// TwinCAT 3 PLC project PLC
// Title: ReMeat003
// Company: Total Control
// Author: Vadim Nagdimaev
// ProjectVersion: 0.0.1
// Description: SLD Line
// ProgramVersion: 3.1.4026.27
// libraries:
//   Tc2_SerialCom, * (Beckhoff Automation GmbH)
//   Tc2_Standard, * (Beckhoff Automation GmbH)
//   Tc2_SUPS, * (Beckhoff Automation GmbH)
//   Tc2_System, * (Beckhoff Automation GmbH)
//   Tc2_Utilities, * (Beckhoff Automation GmbH)
//   Tc3_Module, * (Beckhoff Automation GmbH)
//   Util, * (System)
//   VisuDialogs, * (System)
//   BASIC,3.31,OSCAT
// project tree:
//   00 Library/00-General/ CheckBounds.TcPOU
//   00 Library/00-General/TimeAndDate/ FUN_DeltaTime.TcPOU (excluded from build), GVL_Time_12.TcGVL, prg_RealClock.TcPOU
//   00 Library/00-General/UserGroup/ E_userGroup.TcDUT, prg_User.TcPOU
//   00 Library/01 Piston/ E_ErrorPiton.TcDUT, E_PistonDefault_CMD.TcDUT, E_Piston_Recipe_State.TcDUT, E_Piston_State.TcDUT, FB_Piston.TcPOU, FB_Piston_U_L.TcPOU, ST_Piston.TcDUT, ST_Piston_SelectionList.TcDUT, ST_Piston_Setting_Param.TcDUT, ST_Piston_U_L.TcDUT, TextList_Piston_Recipe_State.TcTLO, TextList_Piston_Recipe_State_CloseOpen.TcTLO, TextList_Piston_Recipe_State_DownUp.TcTLO, TextList_Piston_Recipe_State_InOut.TcTLO, TextList_Piston_Recipe_State_OnOff.TcTLO, TextList_Piston_Recipe_State_OpenClose.TcTLO, TextList_Piston_Recipe_State_UpDown.TcTLO
//   00 Library/01 Piston/VISU/ vis_Piston_Control1.TcVIS, vis_Piston_Control1_Compact.TcVIS, vis_Piston_Control2_CloseOpen.TcVIS, vis_Piston_Control2_OpenClose.TcVIS, vis_Piston_Select.TcVIS (excluded from build), vis_Piston_Select_1.TcVIS (excluded from build), vis_Piston_Setting_Table.TcVIS, vis_Piston_Times.TcVIS
//   00 Library/02 Pump/02.1 Dosing Pump/ FB_DosingPump.TcPOU
//   00 Library/02 Pump/ ControlWordStruct.TcDUT, FB_Pump.TcPOU, StatusWordStruct.TcDUT, ST_Pump.TcDUT
//   00 Library/03 SFC/ FB_SFC_Cycle.TcPOU, FB_SFC_Template.TcPOU, ITF_FB_SFC_Cycle.TcIO, ST_SFC.TcDUT, vis_Cycle_Control.TcVIS, vis_Cycle_Control_1.TcVIS, vis_Cycle_Panel.TcVIS
//   00 Library/04 Recipe/ E_Recipe_Root_Folder.TcDUT, FB_Recipe.TcPOU, FB_Recipe_Vizu.TcVIS, GVL_Recipe.TcGVL, ST_Recipe.TcDUT, TextList_RecipeRootFolder.TcTLO
//   00 Library/04 Recipe/OLD/ prg_RecipeManager.TcPOU, vis_RecipeControl_v01.TcVIS, vis_RecipeTest.TcVIS
//   00 Library/04-Messages/DUTs/Errors/ E_ErrorFormat.TcDUT, ST_Error.TcDUT, ST_Mess_Logger.TcDUT
//   00 Library/04-Messages/DUTs/ stMessageFormat.TcDUT
//   00 Library/04-Messages/ FB_PrintErrMessageByID.TcPOU, FB_PrintErrMessageByID_SFC_Cycle.TcPOU, FB_PrintErrMessageByID_ST_Cycle.TcPOU, FUN_Write_Line_To_History.TcPOU, F_iFB_Num_sFB_Num.TcPOU, GVL_CycleMessages.TcGVL
//   00 Library/05 Safety/ FB_TwinSAFE.TcPOU, GVL_Safety.TcGVL, prg_Safety.TcPOU, ST_ES_PB.TcDUT, ST_SafeOut_PlcIn.TcDUT, ST_SafeIn_PlcOut.TcDUT, Vis_ES_PB.TcVIS
//   00 Library/05 Safety/TwinSAFE/ e_DualChanal.TcDUT, TwinSafeOut_PlcIn.TcDUT, TwinSafeIn_PlcOut.TcDUT
//   00 Library/06-Visu/ ImagePool.TcIPO (not stored), Sensor.TcVIS
//   00 Library/07 Errors/ E_Error_Active_Module.TcDUT, E_OwnerDevice.TcDUT, FB_Error_Handle.TcPOU, ST_DeviceErrorHandeling.TcDUT, vis_Device_Error.TcVIS
//   00 Library/07-Mode/ E_BuzzerMode.TcDUT, E_LightTowerState.TcDUT, E_OperationButtons.TcDUT, E_WorkingMode.TcDUT, FB_ModeSelect.TcPOU, FB_Operation.TcPOU, ST_Mode.TcDUT, ST_OperationButtons.TcDUT
//   00 Library/07-Mode/Visu/ Mode_Select.TcVIS, Mode_Select_1.TcVIS, OperationButtons.TcVIS, OperationButtons_1.TcVIS, OperationButton_Stop.TcVIS, Vis_PauseHistory.TcVIS
//   00 Library/10 Utils/DutyCycle/ FB_DutyCycle.TcPOU, vis_FB_DutyCycle.TcVIS, vis_FB_DutyCycle_Master.TcVIS
//   00 Library/10 Utils/ FB_MovingAverage.TcPOU, FB_Hysteresis_REAL.TcPOU, fun_LrealToString.TcPOU, fun_Real_SecondsToTime.TcPOU, F_TimeRatio.TcPOU, TONR.TcPOU
//   00 Library/11 HMI/ E_Led_Color.TcDUT, g_HMI.TcGVL, ST_MixProof_state.TcDUT
//   00 Library/12 Analog Sensor/ E_ASensor_State.TcTLEO, FB_AnalogSensor.TcPOU, ST_AnalogSensor.TcDUT
//   00 Library/13 Process Control/ FB_ProcessControl.TcPOU, ST_ProcessControl.TcDUT
//   00 Library/30 IO/ FB_ScaleFactor.TcPOU, ST_EL3xx8.TcDUT, ST_EL18x9.TcDUT, ST_EL1918_TwinSafe.TcDUT, ST_EL28x9.TcDUT, ST_EL2904.TcDUT, ST_EL3xx4.TcDUT, ST_EL4xx8.TcDUT, ST_Nidec.TcDUT, ST_TwinSAFE.TcDUT, ST_VTUG.TcDUT
//   00 Library/HeatExchenger/ FB_HeatExchanger.TcPOU, ST_HeatExchanger.TcDUT
//   00 Library/Sensors/ E_Tank_Level.TcDUT, FB_TankSensors.TcPOU, ST_AnalogSignal.TcDUT, ST_Tank_Level.TcDUT
//   01 Instance/00-General/ Global_Constant.TcGVL, Global_Persistent.TcGVL, VersionDescription.TcGVL
//   01 Instance/01 Piston/ E_Pis_Name.TcDUT, g_Piston.TcGVL, prg_Piston.TcPOU
//   01 Instance/02 Pump/ E_Pump_List.TcDUT, g_Pump.TcGVL
//   01 Instance/03 SFC/ g_SFC.TcGVL
//   01 Instance/04 Recipe/ E_Recipe_Name.TcDUT, PlcTask_Recipe.TcTTO, prg_Call_Recipe_Slow.TcPOU, Vis_Recipe_Tab.TcVIS
//   01 Instance/04-Messages/ ERROR_BUFFER.TcVIS, ERROR_HISTORY.TcVIS (excluded from build), Error_List.TcGVL, ERROR_Tab.TcVIS, ERROR_Tab_1.TcVIS, Prg_Filter_Messages.TcPOU, prg_MessageManager.TcPOU, prg_Messages.TcPOU, vis_Error_Act.TcVIS, vis_Error_History.TcVIS, vis_Error_Search.TcVIS
//   01 Instance/06-Visu/ ERRORS_OPER_16_9.TcVIS, ES_INT_OPER_16_9.TcVIS, g_Common.TcGVL, Recipe_16_9.TcVIS
//   01 Instance/06-Visu/Template16-9/ TEMP16_9_00.TcVIS, TEMP16_9_00_1.TcVIS, TEMP16_9_00_Content.TcVIS
//   01 Instance/07-Mode/ E_LightTower_Type.TcDUT, E_ModeZone.TcDUT, E_SkidZone.TcDUT, FB_LightTower.TcPOU, FB_LightTower_Control.TcPOU, GVL_OperMode.TcGVL, prg_Call_OpMode.TcPOU, prg_HMI_OperationLock.TcPOU, prg_LightTower.TcPOU, Vis_LightTower.TcVIS, Vis_LightTower_1.TcVIS, viz_HMI_LockIndex.TcVIS, viz_HMI_Piston.TcVIS
//   01 Instance/12 Analog Sensor/ E_ASense_Name.TcTLEO, g_AnalogSensor.TcGVL
//   01 Instance/13 Process Control/ E_ProcessControl_Name.TcDUT, g_ProcControl.TcGVL
//   03 Project/00 -Initialise/ prg_Initialise.TcPOU (excluded from build)
//   03 Project/23 CIP/ E_Tank_Name.TcTLEO, E_CIP_Client_Command.TcDUT, E_CIP_Client_Selector.TcDUT, E_CIP_DashStage.TcDUT, E_CIP_DashStage_List.TcDUT, E_CIP_Mode.TcDUT, E_CIP_Return.TcDUT, E_CIP_Source.TcDUT, E_CIP_TankList.TcDUT, E_CIP_Type.TcDUT, E_CIP_Usage.TcDUT, FB_CIP.TcPOU, FB_CIP_Client.TcPOU, FB_CIP_Source.TcPOU, FB_CIP_Return.TcPOU, ST_CIP_Param.TcDUT, str_ConcParam.TcDUT, ST_CIP_Request.TcDUT, TextList_CIP_Clients.TcTLO, TextList_CIP_Type.TcTLO, vis_CIP.TcVIS, vis_CIP_ReqBuffer.TcVIS
//   03 Project/21 Data/ E_Element_State_Long.TcDUT
//   03 Project/30 IO/ gIO.TcGVL
//   03 Project/31 AnybusCommunication/ E_Anybus_Alarm.TcDUT, E_Anybus_ClientType.TcDUT, E_Anybus_Media.TcDUT, E_Anybus_RecipeType.TcDUT, E_Anybus_Request.TcDUT, E_Sim_Fault.TcDUT, E_Sim_Mode.TcDUT, FB_Anybus_Interface.TcPOU, FB_CIP_Siemens.TcPOU, FB_Siemens_Sim.TcPOU, ST_Sim_Client.TcDUT, vis_SiemensSim.TcVIS, g_Anybus.TcGVL, ST_Anybus_Inputs.TcDUT, ST_Anybus_Outputs.TcDUT
//   03 Project/ g_Data.TcGVL, vis_Main.TcVIS
//   / GlobalTextList.TcGTLO, PlcTask.TcTTO, RecipeManager.TcRMO (not stored)
//   POUs/ MAIN.TcPOU
// real-time tasks:
//   TASK PlcTask: cycle T#10ms, priority 20, ADS port 350
//   TASK PlcTask_Recipe: cycle T#300ms, priority 14, ADS port 351
//   TASK VISU_TASK: cycle T#200000us, priority 30, ADS port 353
// I/O:
//   DEVICE Device 1 (EtherCAT), AmsNetId 0.0.0.0.2.1
//     BoxTriblrnderBig [EK1200-5000 EtherCAT Power supply (2A E-Bus)]
//       SDI_05 (EL1904) [EL1904, 4 Ch. Safety Input 24V, TwinSAFE]
//         modules: Module 1 (FSOES)
//       SDO_03 (EL2904) [EL2904, 4 Ch. Safety Output 24V, 0.5A, TwinSAFE]
//         modules: Module 1 (FSOES), Module 2 (DO)
//       DI_19 (EL1809) [EL1809 16Ch. Dig. Input 24V, 3ms]
//       DO_11 (EL2809) [EL2809 16Ch. Dig. Output 24V, 0.5A]
//       Term 41 (EL9011) [EL9011 End Terminal]
//   DEVICE Device 2 (EtherCAT), AmsNetId 0.0.0.0.7.1
//     Box 2 (CU1128) [CU1128 6x EtherCAT junction]
//       Box 40 (Anybus Communicator) [Anybus Communicator]
//       BOX_CIP [EK1100 EtherCAT Coupler (2A E-Bus)]
//         SDI_01 (EL1918) [EL1918, 8Ch. Safety Input 24V, TwinSAFE]
//           modules: Module 2 (FSLOGIC)
//         SDI_02 (EL1918) [EL1918, 8Ch. Safety Input 24V, TwinSAFE]
//           modules: Module 1 (FSOE), Module 2 (FSLOGIC)
//         SDO_01 (EL2904) [EL2904, 4 Ch. Safety Output 24V, 0.5A, TwinSAFE]
//           modules: Module 1 (FSOES), Module 2 (DO)
//         DI_01 (EL1809) [EL1809 16Ch. Dig. Input 24V, 3ms]
//         DI_03 (EL1809) [EL1809 16Ch. Dig. Input 24V, 3ms]
//         DI_04 (EL1809) [EL1809 16Ch. Dig. Input 24V, 3ms]
//         DI_05 (EL1809) [EL1809 16Ch. Dig. Input 24V, 3ms]
//         DI_06 (EL1809) [EL1809 16Ch. Dig. Input 24V, 3ms]
//         DO_01 (EL2809) [EL2809 16Ch. Dig. Output 24V, 0.5A]
//         AI_01 (EL3058) [EL3058 8Ch. Ana. Input 4-20mA]
//         AI_02 (EL3058) [EL3058 8Ch. Ana. Input 4-20mA]
//         AO_01 (EL4022) [EL4022 2Ch. Ana. Output 4-20mA, 12bit]
//         Term 103 (EL9011) [EL9011 End Terminal]
//       Box CIP (CTEU-EtherCAT Modular) [CTEU-EtherCAT Fieldbus modular]
//         modules: Module 1 (VAEM-L1-S-24-PT [48DO])
//       Pump CIP (Commander C200 Open Loop) [Commander C200 Open Loop]
//       Box 3 (CU1128-B) [CU1128 6x EtherCAT junction - Dev A]
//         Pump TriBlender (Commander C200 Open Loop) [Commander C200 Open Loop] (disabled)
//       Box 4 (CU1128-C) [CU1128 6x EtherCAT junction - Dev B]
// variable links:
//   Device 1 (EtherCAT) <-> Device 2 (EtherCAT)/Box 2 (CU1128)/BOX_CIP/SDI_01 (EL1918)
//     BoxTriblrnderBig/SDI_05 (EL1904)/Module 1 (FSOES)/RxPDO/FSOE <-> ConnectionInputs/Message_47 TxPDO
//     BoxTriblrnderBig/SDI_05 (EL1904)/Module 1 (FSOES)/TxPDO/FSOE <-> ConnectionOutputs/Message_47 RxPDO
//     BoxTriblrnderBig/SDO_03 (EL2904)/Module 1 (FSOES)/RxPDO/FSOE <-> ConnectionInputs/Message_32 TxPDO
//     BoxTriblrnderBig/SDO_03 (EL2904)/Module 1 (FSOES)/TxPDO/FSOE <-> ConnectionOutputs/Message_32 RxPDO
//   Device 2 (EtherCAT) <-> Device 2 (EtherCAT)/Box 2 (CU1128)/BOX_CIP/SDI_02 (EL1918)
//     Box 2 (CU1128)/BOX_CIP/SDI_01 (EL1918)/ConnectionInputs/Message_10 TxPDO <-> Module 1 (FSOE)/FSoE Outputs/FSOE
//     Box 2 (CU1128)/BOX_CIP/SDI_01 (EL1918)/ConnectionOutputs/Message_10 RxPDO <-> Module 1 (FSOE)/FSoE Inputs/FSOE
//   Device 2 (EtherCAT) <-> Device 2 (EtherCAT)/Box 2 (CU1128)/BOX_CIP/SDO_01 (EL2904)
//     Box 2 (CU1128)/BOX_CIP/SDI_01 (EL1918)/ConnectionInputs/Message_11 TxPDO <-> Module 1 (FSOES)/RxPDO/FSOE
//     Box 2 (CU1128)/BOX_CIP/SDI_01 (EL1918)/ConnectionOutputs/Message_11 RxPDO <-> Module 1 (FSOES)/TxPDO/FSOE
//   PLC/PLC Instance <-> Device 1 (EtherCAT)/BoxTriblrnderBig/DI_19 (EL1809)
//     PlcTask Inputs/gIO.i_EL[19]/i_ch{1..16} <-> Channel {1..16}/Input  (16 links)
//   PLC/PLC Instance <-> Device 1 (EtherCAT)/BoxTriblrnderBig/DO_11 (EL2809)
//     PlcTask Outputs/gIO.q_EL[11]/q_ch{1..16} <-> Channel {1..16}/Output  (16 links)
//   PLC/PLC Instance <-> Device 2 (EtherCAT)/Box 2 (CU1128)/BOX_CIP/AI_01 (EL3058)
//     PlcTask Inputs/gIO.ai_EL[1]/ch{1..8} <-> AI Standard Channel {1..8}/Value  (8 links)
//   PLC/PLC Instance <-> Device 2 (EtherCAT)/Box 2 (CU1128)/BOX_CIP/AI_02 (EL3058)
//     PlcTask Inputs/gIO.ai_EL[2]/ch{1..8} <-> AI Standard Channel {1..8}/Value  (8 links)
//   PLC/PLC Instance <-> Device 2 (EtherCAT)/Box 2 (CU1128)/BOX_CIP/AO_01 (EL4022)
//     PlcTask Outputs/gIO.aq_EL[1]/ch1 <-> AO Outputs Channel 1/Analog output
//     PlcTask Outputs/gIO.aq_EL[1]/ch2 <-> AO Outputs Channel 2/Analog output
//   PLC/PLC Instance <-> Device 2 (EtherCAT)/Box 2 (CU1128)/BOX_CIP/DI_01 (EL1809)
//     PlcTask Inputs/gIO.i_EL[1]/i_ch{1..16} <-> Channel {1..16}/Input  (16 links)
//   PLC/PLC Instance <-> Device 2 (EtherCAT)/Box 2 (CU1128)/BOX_CIP/DI_03 (EL1809)
//     PlcTask Inputs/gIO.i_EL[3]/i_ch{1..16} <-> Channel {1..16}/Input  (16 links)
//   PLC/PLC Instance <-> Device 2 (EtherCAT)/Box 2 (CU1128)/BOX_CIP/DI_04 (EL1809)
//     PlcTask Inputs/gIO.i_EL[4]/i_ch{1..16} <-> Channel {1..16}/Input  (16 links)
//   PLC/PLC Instance <-> Device 2 (EtherCAT)/Box 2 (CU1128)/BOX_CIP/DI_05 (EL1809)
//     PlcTask Inputs/gIO.i_EL[5]/i_ch{1..16} <-> Channel {1..16}/Input  (16 links)
//   PLC/PLC Instance <-> Device 2 (EtherCAT)/Box 2 (CU1128)/BOX_CIP/DI_06 (EL1809)
//     PlcTask Inputs/gIO.i_EL[6]/i_ch{1..16} <-> Channel {1..16}/Input  (16 links)
//   PLC/PLC Instance <-> Device 2 (EtherCAT)/Box 2 (CU1128)/BOX_CIP/DO_01 (EL2809)
//     PlcTask Outputs/gIO.q_EL[1]/q_ch{1..16} <-> Channel {1..16}/Output  (16 links)
//   PLC/PLC Instance <-> Device 2 (EtherCAT)/Box 2 (CU1128)/BOX_CIP/SDI_01 (EL1918)
//     PlcTask Inputs/gIO.arSafe[1].TSafeIn/COM_Err <-> StandardInputs/Standard Out Var 24
//     PlcTask Inputs/gIO.arSafe[1].TSafeIn/FB_Err <-> StandardInputs/Standard Out Var 23
//     PlcTask Inputs/gIO.arSafe[1].TSafeIn/InRun <-> StandardInputs/Standard Out Var 22
//     PlcTask Inputs/gIO.arSafe[1].TSafeIn/Other_Err <-> StandardInputs/Standard Out Var 26
//     PlcTask Inputs/gIO.arSafe[1].stSafetyIn/ES1_PB_State <-> StandardInputs/Standard Out Var 20
//     PlcTask Inputs/gIO.arSafe[1].stSafetyIn/ES2_PB_State <-> StandardInputs/Standard Out Var 40
//     PlcTask Inputs/gIO.arSafe[1].stSafetyIn/ES4_PB_State <-> StandardInputs/Standard Out Var 42
//     PlcTask Inputs/gIO.arSafe[1].stSafetyIn/ES1_State <-> StandardInputs/Standard Out Var 21
//     PlcTask Inputs/gIO.arSafe[1].stSafetyIn/ES2_State <-> StandardInputs/Standard Out Var 38
//     PlcTask Inputs/gIO.arSafe[1].stSafetyIn/ES3_State <-> StandardInputs/Standard Out Var 37
//     PlcTask Inputs/gIO.arSafe[1].stSafetyIn/ES4_State <-> StandardInputs/Standard Out Var 39
//     PlcTask Inputs/gIO.arSafe[1].stSafetyIn/ES3_PB1_State <-> StandardInputs/Standard Out Var 41
//     PlcTask Inputs/gIO.arSafe[1].stSafetyIn/ES3_PB2_State <-> StandardInputs/Standard Out Var 49
//     PlcTask Inputs/gIO.arSafe[1].stSafetyIn/TankLocked_CIP_T{91..94} <-> StandardInputs/Standard Out Var {13..16}  (4 links)
//     PlcTask Inputs/gIO.arSafe[1].stSafetyIn/TankLocked_Color_T3 <-> StandardInputs/Standard Out Var 45
//     PlcTask Inputs/gIO.arSafe[1].stSafetyIn/TankLocked_Color_T4 <-> StandardInputs/Standard Out Var 46
//     PlcTask Inputs/gIO.arSafe[1].stSafetyIn/TankLocked_Marinade_T1 <-> StandardInputs/Standard Out Var 43
//     PlcTask Inputs/gIO.arSafe[1].stSafetyIn/TankLocked_Marinade_T2 <-> StandardInputs/Standard Out Var 44
//     PlcTask Outputs/gIO.arSafe[1].TSafeOut/ErrACK <-> StandardOutputs/Standard In Var 1
//     PlcTask Outputs/gIO.arSafe[1].TSafeOut/RUN <-> StandardOutputs/Standard In Var 2
//     PlcTask Outputs/gIO.arSafe[1].stSafetyOut/ES{1..4}_HMI_PB_Button <-> StandardOutputs/Standard In Var {50..53}  (4 links)
//     PlcTask Outputs/gIO.arSafe[1].stSafetyOut/ES1_PB_Restart <-> StandardOutputs/Standard In Var 28
//     PlcTask Outputs/gIO.arSafe[1].stSafetyOut/ES2_PB_Restart <-> StandardOutputs/Standard In Var 33
//     PlcTask Outputs/gIO.arSafe[1].stSafetyOut/ES3_PB_Restart <-> StandardOutputs/Standard In Var 34
//     PlcTask Outputs/gIO.arSafe[1].stSafetyOut/ES4_PB_Restart <-> StandardOutputs/Standard In Var 35
//   PLC/PLC Instance <-> Device 2 (EtherCAT)/Box 2 (CU1128)/Box 3 (CU1128-B)/Pump TriBlender (Commander C200 Open Loop)
//     PlcTask Inputs/gIO.Nidec[6].StatusWord <-> Transmit PDO Mapping 6/Status word
//     PlcTask Inputs/gIO.Nidec[6].actVelocity <-> Transmit PDO Mapping 6/vl velocity actual value
//     PlcTask Outputs/gIO.Nidec[6].ControlWord <-> Receive PDO Mapping 6/Control word
//     PlcTask Outputs/gIO.Nidec[6].targetVelocity <-> Receive PDO Mapping 6/vl target velocity
//   PLC/PLC Instance <-> Device 2 (EtherCAT)/Box 2 (CU1128)/Box 40 (Anybus Communicator)
//     PlcTask Inputs/gIO.Anybus_Inputs_Raw <-> Transmit PDO Mapping/Input byte 0001
//     PlcTask Inputs/gIO.Anybus_Inputs_Raw @bit 8 <-> Transmit PDO Mapping/Input byte 0002
//     PlcTask Inputs/gIO.Anybus_Inputs_Raw @bit 16 <-> Transmit PDO Mapping/Input byte 0003
//     PlcTask Inputs/gIO.Anybus_Inputs_Raw @bit 24 <-> Transmit PDO Mapping/Input byte 0004
//     PlcTask Inputs/gIO.Anybus_Inputs_Raw @bit 32 <-> Transmit PDO Mapping/Input byte 0005
//     PlcTask Inputs/gIO.Anybus_Inputs_Raw @bit 40 <-> Transmit PDO Mapping/Input byte 0006
//     PlcTask Inputs/gIO.Anybus_Inputs_Raw @bit 48 <-> Transmit PDO Mapping/Input byte 0007
//     PlcTask Inputs/gIO.Anybus_Inputs_Raw @bit 56 <-> Transmit PDO Mapping/Input byte 0008
//     PlcTask Inputs/gIO.Anybus_Inputs_Raw @bit 64 <-> Transmit PDO Mapping/Input byte 0009
//     PlcTask Inputs/gIO.Anybus_Inputs_Raw @bit 72 <-> Transmit PDO Mapping/Input byte 0010
//     PlcTask Inputs/gIO.Anybus_Inputs_Raw @bit 80 <-> Transmit PDO Mapping/Input byte 0011
//     PlcTask Inputs/gIO.Anybus_Inputs_Raw @bit 88 <-> Transmit PDO Mapping/Input byte 0012
//     PlcTask Inputs/gIO.Anybus_Inputs_Raw @bit 96 <-> Transmit PDO Mapping/Input byte 0013
//     PlcTask Inputs/gIO.Anybus_Inputs_Raw @bit 104 <-> Transmit PDO Mapping/Input byte 0014
//     PlcTask Inputs/gIO.Anybus_Inputs_Raw @bit 112 <-> Transmit PDO Mapping/Input byte 0015
//     PlcTask Inputs/gIO.Anybus_Inputs_Raw @bit 120 <-> Transmit PDO Mapping/Input byte 0016
//     PlcTask Inputs/gIO.Anybus_Inputs_Raw @bit 128 <-> Transmit PDO Mapping/Input byte 0017
//     PlcTask Inputs/gIO.Anybus_Inputs_Raw @bit 136 <-> Transmit PDO Mapping/Input byte 0018
//     PlcTask Inputs/gIO.Anybus_Inputs_Raw @bit 144 <-> Transmit PDO Mapping/Input byte 0019
//     PlcTask Inputs/gIO.Anybus_Inputs_Raw @bit 152 <-> Transmit PDO Mapping/Input byte 0020
//     PlcTask Inputs/gIO.Anybus_Inputs_Raw @bit 160 <-> Transmit PDO Mapping/Input byte 0021
//     PlcTask Inputs/gIO.Anybus_Inputs_Raw @bit 168 <-> Transmit PDO Mapping/Input byte 0022
//     PlcTask Inputs/gIO.Anybus_Inputs_Raw @bit 176 <-> Transmit PDO Mapping/Input byte 0023
//     PlcTask Inputs/gIO.Anybus_Inputs_Raw @bit 184 <-> Transmit PDO Mapping/Input byte 0024
//     PlcTask Inputs/gIO.Anybus_Inputs_Raw @bit 192 <-> Transmit PDO Mapping/Input byte 0025
//     PlcTask Inputs/gIO.Anybus_Inputs_Raw @bit 200 <-> Transmit PDO Mapping/Input byte 0026
//     PlcTask Inputs/gIO.Anybus_Inputs_Raw @bit 208 <-> Transmit PDO Mapping/Input byte 0027
//     PlcTask Inputs/gIO.Anybus_Inputs_Raw @bit 216 <-> Transmit PDO Mapping/Input byte 0028
//     PlcTask Inputs/gIO.Anybus_Inputs_Raw @bit 224 <-> Transmit PDO Mapping/Input byte 0029
//     PlcTask Inputs/gIO.Anybus_Inputs_Raw @bit 232 <-> Transmit PDO Mapping/Input byte 0030
//     PlcTask Inputs/gIO.Anybus_Inputs_Raw @bit 240 <-> Transmit PDO Mapping/Input byte 0031
//     PlcTask Inputs/gIO.Anybus_Inputs_Raw @bit 248 <-> Transmit PDO Mapping/Input byte 0032
//     PlcTask Inputs/gIO.Anybus_Inputs_Raw @bit 256 <-> Transmit PDO Mapping/Input byte 0033
//     PlcTask Inputs/gIO.Anybus_Inputs_Raw @bit 264 <-> Transmit PDO Mapping/Input byte 0034
//     PlcTask Inputs/gIO.Anybus_Inputs_Raw @bit 272 <-> Transmit PDO Mapping/Input byte 0035
//     PlcTask Inputs/gIO.Anybus_Inputs_Raw @bit 280 <-> Transmit PDO Mapping/Input byte 0036
//     PlcTask Inputs/gIO.Anybus_Inputs_Raw @bit 288 <-> Transmit PDO Mapping/Input byte 0037
//     PlcTask Inputs/gIO.Anybus_Inputs_Raw @bit 296 <-> Transmit PDO Mapping/Input byte 0038
//     PlcTask Inputs/gIO.Anybus_Inputs_Raw @bit 304 <-> Transmit PDO Mapping/Input byte 0039
//     PlcTask Inputs/gIO.Anybus_Inputs_Raw @bit 312 <-> Transmit PDO Mapping/Input byte 0040
//     PlcTask Inputs/gIO.Anybus_Inputs_Raw @bit 320 <-> Transmit PDO Mapping/Input byte 0041
//     PlcTask Inputs/gIO.Anybus_Inputs_Raw @bit 328 <-> Transmit PDO Mapping/Input byte 0042
//     PlcTask Inputs/gIO.Anybus_Inputs_Raw @bit 336 <-> Transmit PDO Mapping/Input byte 0043
//     PlcTask Inputs/gIO.Anybus_Inputs_Raw @bit 344 <-> Transmit PDO Mapping/Input byte 0044
//     PlcTask Inputs/gIO.Anybus_Inputs_Raw @bit 352 <-> Transmit PDO Mapping/Input byte 0045
//     PlcTask Inputs/gIO.Anybus_Inputs_Raw @bit 360 <-> Transmit PDO Mapping/Input byte 0046
//     PlcTask Inputs/gIO.Anybus_Inputs_Raw @bit 368 <-> Transmit PDO Mapping/Input byte 0047
//     PlcTask Inputs/gIO.Anybus_Inputs_Raw @bit 376 <-> Transmit PDO Mapping/Input byte 0048
//     PlcTask Inputs/gIO.Anybus_Inputs_Raw @bit 384 <-> Transmit PDO Mapping/Input byte 0049
//     PlcTask Inputs/gIO.Anybus_Inputs_Raw @bit 392 <-> Transmit PDO Mapping/Input byte 0050
//     PlcTask Inputs/gIO.Anybus_Inputs_Raw @bit 400 <-> Transmit PDO Mapping/Input byte 0051
//     PlcTask Inputs/gIO.Anybus_Inputs_Raw @bit 408 <-> Transmit PDO Mapping/Input byte 0052
//     PlcTask Inputs/gIO.Anybus_Inputs_Raw @bit 416 <-> Transmit PDO Mapping/Input byte 0053
//     PlcTask Inputs/gIO.Anybus_Inputs_Raw @bit 424 <-> Transmit PDO Mapping/Input byte 0054
//     PlcTask Inputs/gIO.Anybus_Inputs_Raw @bit 432 <-> Transmit PDO Mapping/Input byte 0055
//     PlcTask Inputs/gIO.Anybus_Inputs_Raw @bit 440 <-> Transmit PDO Mapping/Input byte 0056
//     PlcTask Inputs/gIO.Anybus_Inputs_Raw @bit 448 <-> Transmit PDO Mapping/Input byte 0057
//     PlcTask Inputs/gIO.Anybus_Inputs_Raw @bit 456 <-> Transmit PDO Mapping/Input byte 0058
//     PlcTask Inputs/gIO.Anybus_Inputs_Raw @bit 464 <-> Transmit PDO Mapping/Input byte 0059
//     PlcTask Inputs/gIO.Anybus_Inputs_Raw @bit 472 <-> Transmit PDO Mapping/Input byte 0060
//     PlcTask Inputs/gIO.Anybus_Inputs_Raw @bit 480 <-> Transmit PDO Mapping/Input byte 0061
//     PlcTask Inputs/gIO.Anybus_Inputs_Raw @bit 488 <-> Transmit PDO Mapping/Input byte 0062
//     PlcTask Inputs/gIO.Anybus_Inputs_Raw @bit 496 <-> Transmit PDO Mapping/Input byte 0063
//     PlcTask Inputs/gIO.Anybus_Inputs_Raw @bit 504 <-> Transmit PDO Mapping/Input byte 0064
//     PlcTask Inputs/gIO.Anybus_Inputs_Raw @bit 512 <-> Transmit PDO Mapping/Input byte 0065
//     PlcTask Inputs/gIO.Anybus_Inputs_Raw @bit 520 <-> Transmit PDO Mapping/Input byte 0066
//     PlcTask Inputs/gIO.Anybus_Inputs_Raw @bit 528 <-> Transmit PDO Mapping/Input byte 0067
//     PlcTask Inputs/gIO.Anybus_Inputs_Raw @bit 536 <-> Transmit PDO Mapping/Input byte 0068
//     PlcTask Inputs/gIO.Anybus_Inputs_Raw @bit 544 <-> Transmit PDO Mapping/Input byte 0069
//     PlcTask Inputs/gIO.Anybus_Inputs_Raw @bit 552 <-> Transmit PDO Mapping/Input byte 0070
//     PlcTask Inputs/gIO.Anybus_Inputs_Raw @bit 560 <-> Transmit PDO Mapping/Input byte 0071
//     PlcTask Inputs/gIO.Anybus_Inputs_Raw @bit 568 <-> Transmit PDO Mapping/Input byte 0072
//     PlcTask Inputs/gIO.Anybus_Inputs_Raw @bit 576 <-> Transmit PDO Mapping/Input byte 0073
//     PlcTask Inputs/gIO.Anybus_Inputs_Raw @bit 584 <-> Transmit PDO Mapping/Input byte 0074
//     PlcTask Inputs/gIO.Anybus_Inputs_Raw @bit 592 <-> Transmit PDO Mapping/Input byte 0075
//     PlcTask Inputs/gIO.Anybus_Inputs_Raw @bit 600 <-> Transmit PDO Mapping/Input byte 0076
//     PlcTask Inputs/gIO.Anybus_Inputs_Raw @bit 608 <-> Transmit PDO Mapping/Input byte 0077
//     PlcTask Inputs/gIO.Anybus_Inputs_Raw @bit 616 <-> Transmit PDO Mapping/Input byte 0078
//     PlcTask Inputs/gIO.Anybus_Inputs_Raw @bit 624 <-> Transmit PDO Mapping/Input byte 0079
//     PlcTask Inputs/gIO.Anybus_Inputs_Raw @bit 632 <-> Transmit PDO Mapping/Input byte 0080
//     PlcTask Inputs/gIO.Anybus_Inputs_Raw @bit 640 <-> Transmit PDO Mapping/Input byte 0081
//     PlcTask Inputs/gIO.Anybus_Inputs_Raw @bit 648 <-> Transmit PDO Mapping/Input byte 0082
//     PlcTask Inputs/gIO.Anybus_Inputs_Raw @bit 656 <-> Transmit PDO Mapping/Input byte 0083
//     PlcTask Inputs/gIO.Anybus_Inputs_Raw @bit 664 <-> Transmit PDO Mapping/Input byte 0084
//     PlcTask Inputs/gIO.Anybus_Inputs_Raw @bit 672 <-> Transmit PDO Mapping/Input byte 0085
//     PlcTask Inputs/gIO.Anybus_Inputs_Raw @bit 680 <-> Transmit PDO Mapping/Input byte 0086
//     PlcTask Inputs/gIO.Anybus_Inputs_Raw @bit 688 <-> Transmit PDO Mapping/Input byte 0087
//     PlcTask Inputs/gIO.Anybus_Inputs_Raw @bit 696 <-> Transmit PDO Mapping/Input byte 0088
//     PlcTask Inputs/gIO.Anybus_Inputs_Raw @bit 704 <-> Transmit PDO Mapping/Input byte 0089
//     PlcTask Inputs/gIO.Anybus_Inputs_Raw @bit 712 <-> Transmit PDO Mapping/Input byte 0090
//     PlcTask Inputs/gIO.Anybus_Inputs_Raw @bit 720 <-> Transmit PDO Mapping/Input byte 0091
//     PlcTask Inputs/gIO.Anybus_Inputs_Raw @bit 728 <-> Transmit PDO Mapping/Input byte 0092
//     PlcTask Inputs/gIO.Anybus_Inputs_Raw @bit 736 <-> Transmit PDO Mapping/Input byte 0093
//     PlcTask Inputs/gIO.Anybus_Inputs_Raw @bit 744 <-> Transmit PDO Mapping/Input byte 0094
//     PlcTask Inputs/gIO.Anybus_Inputs_Raw @bit 752 <-> Transmit PDO Mapping/Input byte 0095
//     PlcTask Inputs/gIO.Anybus_Inputs_Raw @bit 760 <-> Transmit PDO Mapping/Input byte 0096
//     PlcTask Inputs/gIO.Anybus_Inputs_Raw @bit 768 <-> Transmit PDO Mapping/Input byte 0097
//     PlcTask Inputs/gIO.Anybus_Inputs_Raw @bit 776 <-> Transmit PDO Mapping/Input byte 0098
//     PlcTask Inputs/gIO.Anybus_Inputs_Raw @bit 784 <-> Transmit PDO Mapping/Input byte 0099
//     PlcTask Inputs/gIO.Anybus_Inputs_Raw @bit 792 <-> Transmit PDO Mapping/Input byte 0100
//     PlcTask Inputs/gIO.Anybus_Inputs_Raw @bit 800 <-> Transmit PDO Mapping/Input byte 0101
//     PlcTask Inputs/gIO.Anybus_Inputs_Raw @bit 808 <-> Transmit PDO Mapping/Input byte 0102
//     PlcTask Inputs/gIO.Anybus_Inputs_Raw @bit 816 <-> Transmit PDO Mapping/Input byte 0103
//     PlcTask Inputs/gIO.Anybus_Inputs_Raw @bit 824 <-> Transmit PDO Mapping/Input byte 0104
//     PlcTask Inputs/gIO.Anybus_Inputs_Raw @bit 832 <-> Transmit PDO Mapping/Input byte 0105
//     PlcTask Inputs/gIO.Anybus_Inputs_Raw @bit 840 <-> Transmit PDO Mapping/Input byte 0106
//     PlcTask Inputs/gIO.Anybus_Inputs_Raw @bit 848 <-> Transmit PDO Mapping/Input byte 0107
//     PlcTask Inputs/gIO.Anybus_Inputs_Raw @bit 856 <-> Transmit PDO Mapping/Input byte 0108
//     PlcTask Inputs/gIO.Anybus_Inputs_Raw @bit 864 <-> Transmit PDO Mapping/Input byte 0109
//     PlcTask Inputs/gIO.Anybus_Inputs_Raw @bit 872 <-> Transmit PDO Mapping/Input byte 0110
//     PlcTask Inputs/gIO.Anybus_Inputs_Raw @bit 880 <-> Transmit PDO Mapping/Input byte 0111
//     PlcTask Inputs/gIO.Anybus_Inputs_Raw @bit 888 <-> Transmit PDO Mapping/Input byte 0112
//     PlcTask Inputs/gIO.Anybus_Inputs_Raw @bit 896 <-> Transmit PDO Mapping/Input byte 0113
//     PlcTask Inputs/gIO.Anybus_Inputs_Raw @bit 904 <-> Transmit PDO Mapping/Input byte 0114
//     PlcTask Inputs/gIO.Anybus_Inputs_Raw @bit 912 <-> Transmit PDO Mapping/Input byte 0115
//     PlcTask Inputs/gIO.Anybus_Inputs_Raw @bit 920 <-> Transmit PDO Mapping/Input byte 0116
//     PlcTask Inputs/gIO.Anybus_Inputs_Raw @bit 928 <-> Transmit PDO Mapping/Input byte 0117
//     PlcTask Inputs/gIO.Anybus_Inputs_Raw @bit 936 <-> Transmit PDO Mapping/Input byte 0118
//     PlcTask Inputs/gIO.Anybus_Inputs_Raw @bit 944 <-> Transmit PDO Mapping/Input byte 0119
//     PlcTask Inputs/gIO.Anybus_Inputs_Raw @bit 952 <-> Transmit PDO Mapping/Input byte 0120
//     PlcTask Inputs/gIO.Anybus_Inputs_Raw @bit 960 <-> Transmit PDO Mapping/Input byte 0121
//     PlcTask Inputs/gIO.Anybus_Inputs_Raw @bit 968 <-> Transmit PDO Mapping/Input byte 0122
//     PlcTask Inputs/gIO.Anybus_Inputs_Raw @bit 976 <-> Transmit PDO Mapping/Input byte 0123
//     PlcTask Inputs/gIO.Anybus_Inputs_Raw @bit 984 <-> Transmit PDO Mapping/Input byte 0124
//     PlcTask Inputs/gIO.Anybus_Inputs_Raw @bit 992 <-> Transmit PDO Mapping/Input byte 0125
//     PlcTask Inputs/gIO.Anybus_Inputs_Raw @bit 1000 <-> Transmit PDO Mapping/Input byte 0126
//     PlcTask Inputs/gIO.Anybus_Inputs_Raw @bit 1008 <-> Transmit PDO Mapping/Input byte 0127
//     PlcTask Inputs/gIO.Anybus_Inputs_Raw @bit 1016 <-> Transmit PDO Mapping/Input byte 0128
//     PlcTask Inputs/gIO.Anybus_WcState <-> WcState/WcState
//     PlcTask Outputs/gIO.Anybus_Outputs_Raw <-> Receive PDO Mapping/Output byte 0001
//     PlcTask Outputs/gIO.Anybus_Outputs_Raw @bit 8 <-> Receive PDO Mapping/Output byte 0002
//     PlcTask Outputs/gIO.Anybus_Outputs_Raw @bit 16 <-> Receive PDO Mapping/Output byte 0003
//     PlcTask Outputs/gIO.Anybus_Outputs_Raw @bit 24 <-> Receive PDO Mapping/Output byte 0004
//     PlcTask Outputs/gIO.Anybus_Outputs_Raw @bit 32 <-> Receive PDO Mapping/Output byte 0005
//     PlcTask Outputs/gIO.Anybus_Outputs_Raw @bit 40 <-> Receive PDO Mapping/Output byte 0006
//     PlcTask Outputs/gIO.Anybus_Outputs_Raw @bit 48 <-> Receive PDO Mapping/Output byte 0007
//     PlcTask Outputs/gIO.Anybus_Outputs_Raw @bit 56 <-> Receive PDO Mapping/Output byte 0008
//     PlcTask Outputs/gIO.Anybus_Outputs_Raw @bit 64 <-> Receive PDO Mapping/Output byte 0009
//     PlcTask Outputs/gIO.Anybus_Outputs_Raw @bit 72 <-> Receive PDO Mapping/Output byte 0010
//     PlcTask Outputs/gIO.Anybus_Outputs_Raw @bit 80 <-> Receive PDO Mapping/Output byte 0011
//     PlcTask Outputs/gIO.Anybus_Outputs_Raw @bit 88 <-> Receive PDO Mapping/Output byte 0012
//     PlcTask Outputs/gIO.Anybus_Outputs_Raw @bit 96 <-> Receive PDO Mapping/Output byte 0013
//     PlcTask Outputs/gIO.Anybus_Outputs_Raw @bit 104 <-> Receive PDO Mapping/Output byte 0014
//     PlcTask Outputs/gIO.Anybus_Outputs_Raw @bit 112 <-> Receive PDO Mapping/Output byte 0015
//     PlcTask Outputs/gIO.Anybus_Outputs_Raw @bit 120 <-> Receive PDO Mapping/Output byte 0016
//     PlcTask Outputs/gIO.Anybus_Outputs_Raw @bit 128 <-> Receive PDO Mapping/Output byte 0017
//     PlcTask Outputs/gIO.Anybus_Outputs_Raw @bit 136 <-> Receive PDO Mapping/Output byte 0018
//     PlcTask Outputs/gIO.Anybus_Outputs_Raw @bit 144 <-> Receive PDO Mapping/Output byte 0019
//     PlcTask Outputs/gIO.Anybus_Outputs_Raw @bit 152 <-> Receive PDO Mapping/Output byte 0020
//     PlcTask Outputs/gIO.Anybus_Outputs_Raw @bit 160 <-> Receive PDO Mapping/Output byte 0021
//     PlcTask Outputs/gIO.Anybus_Outputs_Raw @bit 168 <-> Receive PDO Mapping/Output byte 0022
//     PlcTask Outputs/gIO.Anybus_Outputs_Raw @bit 176 <-> Receive PDO Mapping/Output byte 0023
//     PlcTask Outputs/gIO.Anybus_Outputs_Raw @bit 184 <-> Receive PDO Mapping/Output byte 0024
//     PlcTask Outputs/gIO.Anybus_Outputs_Raw @bit 192 <-> Receive PDO Mapping/Output byte 0025
//     PlcTask Outputs/gIO.Anybus_Outputs_Raw @bit 200 <-> Receive PDO Mapping/Output byte 0026
//     PlcTask Outputs/gIO.Anybus_Outputs_Raw @bit 208 <-> Receive PDO Mapping/Output byte 0027
//     PlcTask Outputs/gIO.Anybus_Outputs_Raw @bit 216 <-> Receive PDO Mapping/Output byte 0028
//     PlcTask Outputs/gIO.Anybus_Outputs_Raw @bit 224 <-> Receive PDO Mapping/Output byte 0029
//     PlcTask Outputs/gIO.Anybus_Outputs_Raw @bit 232 <-> Receive PDO Mapping/Output byte 0030
//     PlcTask Outputs/gIO.Anybus_Outputs_Raw @bit 240 <-> Receive PDO Mapping/Output byte 0031
//     PlcTask Outputs/gIO.Anybus_Outputs_Raw @bit 248 <-> Receive PDO Mapping/Output byte 0032
//     PlcTask Outputs/gIO.Anybus_Outputs_Raw @bit 256 <-> Receive PDO Mapping/Output byte 0033
//     PlcTask Outputs/gIO.Anybus_Outputs_Raw @bit 264 <-> Receive PDO Mapping/Output byte 0034
//     PlcTask Outputs/gIO.Anybus_Outputs_Raw @bit 272 <-> Receive PDO Mapping/Output byte 0035
//     PlcTask Outputs/gIO.Anybus_Outputs_Raw @bit 280 <-> Receive PDO Mapping/Output byte 0036
//     PlcTask Outputs/gIO.Anybus_Outputs_Raw @bit 288 <-> Receive PDO Mapping/Output byte 0037
//     PlcTask Outputs/gIO.Anybus_Outputs_Raw @bit 296 <-> Receive PDO Mapping/Output byte 0038
//     PlcTask Outputs/gIO.Anybus_Outputs_Raw @bit 304 <-> Receive PDO Mapping/Output byte 0039
//     PlcTask Outputs/gIO.Anybus_Outputs_Raw @bit 312 <-> Receive PDO Mapping/Output byte 0040
//     PlcTask Outputs/gIO.Anybus_Outputs_Raw @bit 320 <-> Receive PDO Mapping/Output byte 0041
//     PlcTask Outputs/gIO.Anybus_Outputs_Raw @bit 328 <-> Receive PDO Mapping/Output byte 0042
//     PlcTask Outputs/gIO.Anybus_Outputs_Raw @bit 336 <-> Receive PDO Mapping/Output byte 0043
//     PlcTask Outputs/gIO.Anybus_Outputs_Raw @bit 344 <-> Receive PDO Mapping/Output byte 0044
//     PlcTask Outputs/gIO.Anybus_Outputs_Raw @bit 352 <-> Receive PDO Mapping/Output byte 0045
//     PlcTask Outputs/gIO.Anybus_Outputs_Raw @bit 360 <-> Receive PDO Mapping/Output byte 0046
//     PlcTask Outputs/gIO.Anybus_Outputs_Raw @bit 368 <-> Receive PDO Mapping/Output byte 0047
//     PlcTask Outputs/gIO.Anybus_Outputs_Raw @bit 376 <-> Receive PDO Mapping/Output byte 0048
//     PlcTask Outputs/gIO.Anybus_Outputs_Raw @bit 384 <-> Receive PDO Mapping/Output byte 0049
//     PlcTask Outputs/gIO.Anybus_Outputs_Raw @bit 392 <-> Receive PDO Mapping/Output byte 0050
//     PlcTask Outputs/gIO.Anybus_Outputs_Raw @bit 400 <-> Receive PDO Mapping/Output byte 0051
//     PlcTask Outputs/gIO.Anybus_Outputs_Raw @bit 408 <-> Receive PDO Mapping/Output byte 0052
//     PlcTask Outputs/gIO.Anybus_Outputs_Raw @bit 416 <-> Receive PDO Mapping/Output byte 0053
//     PlcTask Outputs/gIO.Anybus_Outputs_Raw @bit 424 <-> Receive PDO Mapping/Output byte 0054
//     PlcTask Outputs/gIO.Anybus_Outputs_Raw @bit 432 <-> Receive PDO Mapping/Output byte 0055
//     PlcTask Outputs/gIO.Anybus_Outputs_Raw @bit 440 <-> Receive PDO Mapping/Output byte 0056
//     PlcTask Outputs/gIO.Anybus_Outputs_Raw @bit 448 <-> Receive PDO Mapping/Output byte 0057
//     PlcTask Outputs/gIO.Anybus_Outputs_Raw @bit 456 <-> Receive PDO Mapping/Output byte 0058
//     PlcTask Outputs/gIO.Anybus_Outputs_Raw @bit 464 <-> Receive PDO Mapping/Output byte 0059
//     PlcTask Outputs/gIO.Anybus_Outputs_Raw @bit 472 <-> Receive PDO Mapping/Output byte 0060
//     PlcTask Outputs/gIO.Anybus_Outputs_Raw @bit 480 <-> Receive PDO Mapping/Output byte 0061
//     PlcTask Outputs/gIO.Anybus_Outputs_Raw @bit 488 <-> Receive PDO Mapping/Output byte 0062
//     PlcTask Outputs/gIO.Anybus_Outputs_Raw @bit 496 <-> Receive PDO Mapping/Output byte 0063
//     PlcTask Outputs/gIO.Anybus_Outputs_Raw @bit 504 <-> Receive PDO Mapping/Output byte 0064
//     PlcTask Outputs/gIO.Anybus_Outputs_Raw @bit 512 <-> Receive PDO Mapping/Output byte 0065
//     PlcTask Outputs/gIO.Anybus_Outputs_Raw @bit 520 <-> Receive PDO Mapping/Output byte 0066
//     PlcTask Outputs/gIO.Anybus_Outputs_Raw @bit 528 <-> Receive PDO Mapping/Output byte 0067
//     PlcTask Outputs/gIO.Anybus_Outputs_Raw @bit 536 <-> Receive PDO Mapping/Output byte 0068
//     PlcTask Outputs/gIO.Anybus_Outputs_Raw @bit 544 <-> Receive PDO Mapping/Output byte 0069
//     PlcTask Outputs/gIO.Anybus_Outputs_Raw @bit 552 <-> Receive PDO Mapping/Output byte 0070
//     PlcTask Outputs/gIO.Anybus_Outputs_Raw @bit 560 <-> Receive PDO Mapping/Output byte 0071
//     PlcTask Outputs/gIO.Anybus_Outputs_Raw @bit 568 <-> Receive PDO Mapping/Output byte 0072
//     PlcTask Outputs/gIO.Anybus_Outputs_Raw @bit 576 <-> Receive PDO Mapping/Output byte 0073
//     PlcTask Outputs/gIO.Anybus_Outputs_Raw @bit 584 <-> Receive PDO Mapping/Output byte 0074
//     PlcTask Outputs/gIO.Anybus_Outputs_Raw @bit 592 <-> Receive PDO Mapping/Output byte 0075
//     PlcTask Outputs/gIO.Anybus_Outputs_Raw @bit 600 <-> Receive PDO Mapping/Output byte 0076
//     PlcTask Outputs/gIO.Anybus_Outputs_Raw @bit 608 <-> Receive PDO Mapping/Output byte 0077
//     PlcTask Outputs/gIO.Anybus_Outputs_Raw @bit 616 <-> Receive PDO Mapping/Output byte 0078
//     PlcTask Outputs/gIO.Anybus_Outputs_Raw @bit 624 <-> Receive PDO Mapping/Output byte 0079
//     PlcTask Outputs/gIO.Anybus_Outputs_Raw @bit 632 <-> Receive PDO Mapping/Output byte 0080
//     PlcTask Outputs/gIO.Anybus_Outputs_Raw @bit 640 <-> Receive PDO Mapping/Output byte 0081
//     PlcTask Outputs/gIO.Anybus_Outputs_Raw @bit 648 <-> Receive PDO Mapping/Output byte 0082
//     PlcTask Outputs/gIO.Anybus_Outputs_Raw @bit 656 <-> Receive PDO Mapping/Output byte 0083
//     PlcTask Outputs/gIO.Anybus_Outputs_Raw @bit 664 <-> Receive PDO Mapping/Output byte 0084
//     PlcTask Outputs/gIO.Anybus_Outputs_Raw @bit 672 <-> Receive PDO Mapping/Output byte 0085
//     PlcTask Outputs/gIO.Anybus_Outputs_Raw @bit 680 <-> Receive PDO Mapping/Output byte 0086
//     PlcTask Outputs/gIO.Anybus_Outputs_Raw @bit 688 <-> Receive PDO Mapping/Output byte 0087
//     PlcTask Outputs/gIO.Anybus_Outputs_Raw @bit 696 <-> Receive PDO Mapping/Output byte 0088
//     PlcTask Outputs/gIO.Anybus_Outputs_Raw @bit 704 <-> Receive PDO Mapping/Output byte 0089
//     PlcTask Outputs/gIO.Anybus_Outputs_Raw @bit 712 <-> Receive PDO Mapping/Output byte 0090
//     PlcTask Outputs/gIO.Anybus_Outputs_Raw @bit 720 <-> Receive PDO Mapping/Output byte 0091
//     PlcTask Outputs/gIO.Anybus_Outputs_Raw @bit 728 <-> Receive PDO Mapping/Output byte 0092
//     PlcTask Outputs/gIO.Anybus_Outputs_Raw @bit 736 <-> Receive PDO Mapping/Output byte 0093
//     PlcTask Outputs/gIO.Anybus_Outputs_Raw @bit 744 <-> Receive PDO Mapping/Output byte 0094
//     PlcTask Outputs/gIO.Anybus_Outputs_Raw @bit 752 <-> Receive PDO Mapping/Output byte 0095
//     PlcTask Outputs/gIO.Anybus_Outputs_Raw @bit 760 <-> Receive PDO Mapping/Output byte 0096
//     PlcTask Outputs/gIO.Anybus_Outputs_Raw @bit 768 <-> Receive PDO Mapping/Output byte 0097
//     PlcTask Outputs/gIO.Anybus_Outputs_Raw @bit 776 <-> Receive PDO Mapping/Output byte 0098
//     PlcTask Outputs/gIO.Anybus_Outputs_Raw @bit 784 <-> Receive PDO Mapping/Output byte 0099
//     PlcTask Outputs/gIO.Anybus_Outputs_Raw @bit 792 <-> Receive PDO Mapping/Output byte 0100
//     PlcTask Outputs/gIO.Anybus_Outputs_Raw @bit 800 <-> Receive PDO Mapping/Output byte 0101
//     PlcTask Outputs/gIO.Anybus_Outputs_Raw @bit 808 <-> Receive PDO Mapping/Output byte 0102
//     PlcTask Outputs/gIO.Anybus_Outputs_Raw @bit 816 <-> Receive PDO Mapping/Output byte 0103
//     PlcTask Outputs/gIO.Anybus_Outputs_Raw @bit 824 <-> Receive PDO Mapping/Output byte 0104
//     PlcTask Outputs/gIO.Anybus_Outputs_Raw @bit 832 <-> Receive PDO Mapping/Output byte 0105
//     PlcTask Outputs/gIO.Anybus_Outputs_Raw @bit 840 <-> Receive PDO Mapping/Output byte 0106
//     PlcTask Outputs/gIO.Anybus_Outputs_Raw @bit 848 <-> Receive PDO Mapping/Output byte 0107
//     PlcTask Outputs/gIO.Anybus_Outputs_Raw @bit 856 <-> Receive PDO Mapping/Output byte 0108
//     PlcTask Outputs/gIO.Anybus_Outputs_Raw @bit 864 <-> Receive PDO Mapping/Output byte 0109
//     PlcTask Outputs/gIO.Anybus_Outputs_Raw @bit 872 <-> Receive PDO Mapping/Output byte 0110
//     PlcTask Outputs/gIO.Anybus_Outputs_Raw @bit 880 <-> Receive PDO Mapping/Output byte 0111
//     PlcTask Outputs/gIO.Anybus_Outputs_Raw @bit 888 <-> Receive PDO Mapping/Output byte 0112
//     PlcTask Outputs/gIO.Anybus_Outputs_Raw @bit 896 <-> Receive PDO Mapping/Output byte 0113
//     PlcTask Outputs/gIO.Anybus_Outputs_Raw @bit 904 <-> Receive PDO Mapping/Output byte 0114
//     PlcTask Outputs/gIO.Anybus_Outputs_Raw @bit 912 <-> Receive PDO Mapping/Output byte 0115
//     PlcTask Outputs/gIO.Anybus_Outputs_Raw @bit 920 <-> Receive PDO Mapping/Output byte 0116
//     PlcTask Outputs/gIO.Anybus_Outputs_Raw @bit 928 <-> Receive PDO Mapping/Output byte 0117
//     PlcTask Outputs/gIO.Anybus_Outputs_Raw @bit 936 <-> Receive PDO Mapping/Output byte 0118
//     PlcTask Outputs/gIO.Anybus_Outputs_Raw @bit 944 <-> Receive PDO Mapping/Output byte 0119
//     PlcTask Outputs/gIO.Anybus_Outputs_Raw @bit 952 <-> Receive PDO Mapping/Output byte 0120
//     PlcTask Outputs/gIO.Anybus_Outputs_Raw @bit 960 <-> Receive PDO Mapping/Output byte 0121
//     PlcTask Outputs/gIO.Anybus_Outputs_Raw @bit 968 <-> Receive PDO Mapping/Output byte 0122
//     PlcTask Outputs/gIO.Anybus_Outputs_Raw @bit 976 <-> Receive PDO Mapping/Output byte 0123
//     PlcTask Outputs/gIO.Anybus_Outputs_Raw @bit 984 <-> Receive PDO Mapping/Output byte 0124
//     PlcTask Outputs/gIO.Anybus_Outputs_Raw @bit 992 <-> Receive PDO Mapping/Output byte 0125
//     PlcTask Outputs/gIO.Anybus_Outputs_Raw @bit 1000 <-> Receive PDO Mapping/Output byte 0126
//     PlcTask Outputs/gIO.Anybus_Outputs_Raw @bit 1008 <-> Receive PDO Mapping/Output byte 0127
//     PlcTask Outputs/gIO.Anybus_Outputs_Raw @bit 1016 <-> Receive PDO Mapping/Output byte 0128
//   PLC/PLC Instance <-> Device 2 (EtherCAT)/Box 2 (CU1128)/Box CIP (CTEU-EtherCAT Modular)
//     PlcTask Outputs/gIO.q_Manifold1[10]/sol_12 <-> Module 1 (VAEM-L1-S-24-PT [48DO])/Outputs/C3 Output[3]
//     PlcTask Outputs/gIO.q_Manifold1[10]/sol_14 <-> Module 1 (VAEM-L1-S-24-PT [48DO])/Outputs/C3 Output[2]
//     PlcTask Outputs/gIO.q_Manifold1[11]/sol_12 <-> Module 1 (VAEM-L1-S-24-PT [48DO])/Outputs/C3 Output[5]
//     PlcTask Outputs/gIO.q_Manifold1[11]/sol_14 <-> Module 1 (VAEM-L1-S-24-PT [48DO])/Outputs/C3 Output[4]
//     PlcTask Outputs/gIO.q_Manifold1[12]/sol_12 <-> Module 1 (VAEM-L1-S-24-PT [48DO])/Outputs/C3 Output[7]
//     PlcTask Outputs/gIO.q_Manifold1[12]/sol_14 <-> Module 1 (VAEM-L1-S-24-PT [48DO])/Outputs/C3 Output[6]
//     PlcTask Outputs/gIO.q_Manifold1[13]/sol_12 <-> Module 1 (VAEM-L1-S-24-PT [48DO])/Outputs/C4 Output[1]
//     PlcTask Outputs/gIO.q_Manifold1[13]/sol_14 <-> Module 1 (VAEM-L1-S-24-PT [48DO])/Outputs/C4 Output[0]
//     PlcTask Outputs/gIO.q_Manifold1[14]/sol_12 <-> Module 1 (VAEM-L1-S-24-PT [48DO])/Outputs/C4 Output[3]
//     PlcTask Outputs/gIO.q_Manifold1[14]/sol_14 <-> Module 1 (VAEM-L1-S-24-PT [48DO])/Outputs/C4 Output[2]
//     PlcTask Outputs/gIO.q_Manifold1[15]/sol_12 <-> Module 1 (VAEM-L1-S-24-PT [48DO])/Outputs/C4 Output[5]
//     PlcTask Outputs/gIO.q_Manifold1[15]/sol_14 <-> Module 1 (VAEM-L1-S-24-PT [48DO])/Outputs/C4 Output[4]
//     PlcTask Outputs/gIO.q_Manifold1[16]/sol_12 <-> Module 1 (VAEM-L1-S-24-PT [48DO])/Outputs/C4 Output[7]
//     PlcTask Outputs/gIO.q_Manifold1[16]/sol_14 <-> Module 1 (VAEM-L1-S-24-PT [48DO])/Outputs/C4 Output[6]
//     PlcTask Outputs/gIO.q_Manifold1[17]/sol_12 <-> Module 1 (VAEM-L1-S-24-PT [48DO])/Outputs/C5 Output[1]
//     PlcTask Outputs/gIO.q_Manifold1[17]/sol_14 <-> Module 1 (VAEM-L1-S-24-PT [48DO])/Outputs/C5 Output[0]
//     PlcTask Outputs/gIO.q_Manifold1[18]/sol_12 <-> Module 1 (VAEM-L1-S-24-PT [48DO])/Outputs/C5 Output[3]
//     PlcTask Outputs/gIO.q_Manifold1[18]/sol_14 <-> Module 1 (VAEM-L1-S-24-PT [48DO])/Outputs/C5 Output[2]
//     PlcTask Outputs/gIO.q_Manifold1[19]/sol_12 <-> Module 1 (VAEM-L1-S-24-PT [48DO])/Outputs/C5 Output[5]
//     PlcTask Outputs/gIO.q_Manifold1[19]/sol_14 <-> Module 1 (VAEM-L1-S-24-PT [48DO])/Outputs/C5 Output[4]
//     PlcTask Outputs/gIO.q_Manifold1[1]/sol_12 <-> Module 1 (VAEM-L1-S-24-PT [48DO])/Outputs/C1 Output[1]
//     PlcTask Outputs/gIO.q_Manifold1[1]/sol_14 <-> Module 1 (VAEM-L1-S-24-PT [48DO])/Outputs/C1 Output[0]
//     PlcTask Outputs/gIO.q_Manifold1[20]/sol_12 <-> Module 1 (VAEM-L1-S-24-PT [48DO])/Outputs/C5 Output[7]
//     PlcTask Outputs/gIO.q_Manifold1[20]/sol_14 <-> Module 1 (VAEM-L1-S-24-PT [48DO])/Outputs/C5 Output[6]
//     PlcTask Outputs/gIO.q_Manifold1[21]/sol_12 <-> Module 1 (VAEM-L1-S-24-PT [48DO])/Outputs/C6 Output[1]
//     PlcTask Outputs/gIO.q_Manifold1[21]/sol_14 <-> Module 1 (VAEM-L1-S-24-PT [48DO])/Outputs/C6 Output[0]
//     PlcTask Outputs/gIO.q_Manifold1[22]/sol_12 <-> Module 1 (VAEM-L1-S-24-PT [48DO])/Outputs/C6 Output[3]
//     PlcTask Outputs/gIO.q_Manifold1[22]/sol_14 <-> Module 1 (VAEM-L1-S-24-PT [48DO])/Outputs/C6 Output[2]
//     PlcTask Outputs/gIO.q_Manifold1[23]/sol_12 <-> Module 1 (VAEM-L1-S-24-PT [48DO])/Outputs/C6 Output[5]
//     PlcTask Outputs/gIO.q_Manifold1[23]/sol_14 <-> Module 1 (VAEM-L1-S-24-PT [48DO])/Outputs/C6 Output[4]
//     PlcTask Outputs/gIO.q_Manifold1[24]/sol_12 <-> Module 1 (VAEM-L1-S-24-PT [48DO])/Outputs/C6 Output[7]
//     PlcTask Outputs/gIO.q_Manifold1[24]/sol_14 <-> Module 1 (VAEM-L1-S-24-PT [48DO])/Outputs/C6 Output[6]
//     PlcTask Outputs/gIO.q_Manifold1[2]/sol_12 <-> Module 1 (VAEM-L1-S-24-PT [48DO])/Outputs/C1 Output[3]
//     PlcTask Outputs/gIO.q_Manifold1[2]/sol_14 <-> Module 1 (VAEM-L1-S-24-PT [48DO])/Outputs/C1 Output[2]
//     PlcTask Outputs/gIO.q_Manifold1[3]/sol_12 <-> Module 1 (VAEM-L1-S-24-PT [48DO])/Outputs/C1 Output[5]
//     PlcTask Outputs/gIO.q_Manifold1[3]/sol_14 <-> Module 1 (VAEM-L1-S-24-PT [48DO])/Outputs/C1 Output[4]
//     PlcTask Outputs/gIO.q_Manifold1[4]/sol_12 <-> Module 1 (VAEM-L1-S-24-PT [48DO])/Outputs/C1 Output[7]
//     PlcTask Outputs/gIO.q_Manifold1[4]/sol_14 <-> Module 1 (VAEM-L1-S-24-PT [48DO])/Outputs/C1 Output[6]
//     PlcTask Outputs/gIO.q_Manifold1[5]/sol_12 <-> Module 1 (VAEM-L1-S-24-PT [48DO])/Outputs/C2 Output[1]
//     PlcTask Outputs/gIO.q_Manifold1[5]/sol_14 <-> Module 1 (VAEM-L1-S-24-PT [48DO])/Outputs/C2 Output[0]
//     PlcTask Outputs/gIO.q_Manifold1[6]/sol_12 <-> Module 1 (VAEM-L1-S-24-PT [48DO])/Outputs/C2 Output[3]
//     PlcTask Outputs/gIO.q_Manifold1[6]/sol_14 <-> Module 1 (VAEM-L1-S-24-PT [48DO])/Outputs/C2 Output[2]
//     PlcTask Outputs/gIO.q_Manifold1[7]/sol_12 <-> Module 1 (VAEM-L1-S-24-PT [48DO])/Outputs/C2 Output[5]
//     PlcTask Outputs/gIO.q_Manifold1[7]/sol_14 <-> Module 1 (VAEM-L1-S-24-PT [48DO])/Outputs/C2 Output[4]
//     PlcTask Outputs/gIO.q_Manifold1[8]/sol_12 <-> Module 1 (VAEM-L1-S-24-PT [48DO])/Outputs/C2 Output[7]
//     PlcTask Outputs/gIO.q_Manifold1[8]/sol_14 <-> Module 1 (VAEM-L1-S-24-PT [48DO])/Outputs/C2 Output[6]
//     PlcTask Outputs/gIO.q_Manifold1[9]/sol_12 <-> Module 1 (VAEM-L1-S-24-PT [48DO])/Outputs/C3 Output[1]
//     PlcTask Outputs/gIO.q_Manifold1[9]/sol_14 <-> Module 1 (VAEM-L1-S-24-PT [48DO])/Outputs/C3 Output[0]
//   PLC/PLC Instance <-> Device 2 (EtherCAT)/Box 2 (CU1128)/Pump CIP (Commander C200 Open Loop)
//     PlcTask Inputs/gIO.Nidec[1].StatusWord <-> Transmit PDO Mapping 6/Status word
//     PlcTask Inputs/gIO.Nidec[1].actVelocity <-> Transmit PDO Mapping 6/vl velocity actual value
//     PlcTask Outputs/gIO.Nidec[1].ControlWord <-> Receive PDO Mapping 6/Control word
//     PlcTask Outputs/gIO.Nidec[1].targetVelocity <-> Receive PDO Mapping 6/vl target velocity

CONFIGURATION PLC
    RESOURCE PLC ON TwinCAT3
        TASK PlcTask_Recipe(INTERVAL := T#300ms, PRIORITY := 14);
        TASK PlcTask(INTERVAL := T#10ms, PRIORITY := 20);
        PROGRAM prg_Call_Recipe_Slow WITH PlcTask_Recipe : prg_Call_Recipe_Slow;
        PROGRAM MAIN WITH PlcTask : MAIN;
    END_RESOURCE
END_CONFIGURATION

// ---- 00 Library/00-General/UserGroup/E_userGroup.TcDUT

TYPE E_userGroup :
(
	Group1:=1,
	Group2:=2,
	Group3:=3,
	Group4:=4
);
END_TYPE

// ---- 00 Library/01 Piston/E_ErrorPiton.TcDUT
{attribute 'qualified_only'}
{attribute 'strict'}
TYPE E_ErrorPiton :
(
	No_piston_error							:=0,
	Wating_for_sensor_open_at_Open_cmd		:=1,
	Wating_for_sensor_close_at_Open_cmd		:=2,
	Wating_for_sensor_close_at_Close_cmd	:=3,
	Wating_for_sensor_open_at_Close_cmd		:=4,
	No_status								:=5,
	No_valve_Operation						:=6,
	Error_not_difined						:=9);
END_TYPE

// ---- 00 Library/01 Piston/E_PistonDefault_CMD.TcDUT
{attribute 'qualified_only'}
{attribute 'strict'}
TYPE E_PistonDefault_CMD :
(
	Close := 0,
	Open,
	Sensors, 		//by actual sensors state
	SensorsClose,	//by actual sensors state, if state wrong close
	SensorsOpen		//by actual sensors state, if state wrong open
);
END_TYPE

// ---- 00 Library/01 Piston/E_Piston_Recipe_State.TcDUT
{attribute 'qualified_only'}
{attribute 'strict'}
TYPE E_Piston_Recipe_State :
(
	NoChanges := 0,
	Act,	// action invert deafult cmd
	Release	// action deafult cmd
);
END_TYPE

// ---- 00 Library/01 Piston/E_Piston_State.TcDUT
{attribute 'qualified_only'}
{attribute 'strict'}
TYPE E_Piston_State :
(
	Init := 0,
	Close,Open,Busy_Close,Busy_Open
);
END_TYPE

// ---- 00 Library/01 Piston/ST_Piston.TcDUT
TYPE ST_Piston :
STRUCT
	req_Open		:BOOL;		(* Auto cycle command, will operate the piston to open, not for HMI usage	*)
	req_Close		:BOOL;		(* Auto cycle command, will operate the piston to close, not for HMI usage	*)
	
	//additional requests for Upper and Lower 
	req_Upper		:	BOOL	;
	req_Lower		:	BOOL	;

	req_OpenMan		:BOOL;		(* Manual command, for HMI, will operate the piston to open	*)
	req_CloseMan	:BOOL;		(* Manual command, for HMI, will operate the piston to close	*)
	req_DefaultPos	:BOOL;		(* Manual command, for HMI, will operate the piston to its default position*)

	b_Enable		: BOOL:=TRUE;(* Piston operation enable,  *)
	b_Reset			: BOOL;		(* The command will reset all commands and cycle state*)
	b_Resume		: BOOL;		(* In case of malfunction the function getting pause state, the command will resume the cycle flow *)
	b_Error			: BOOL;
	b_Exist			: BOOL;		(*FB_Piston executed - avalable for visu*)
	b_InterLock		: BOOL 	:=TRUE;
	b_InterLock_Open		: BOOL 	:=TRUE;
	b_InterLock_Close		: BOOL 	:=TRUE;
	b_DeactivateMan	: BOOL;


	// Status
	st_Open			: BOOL	:=FALSE;	(* Piston state open	*)
	st_Close		: BOOL	:=FALSE;	(* Piston state close	*)	
	st_Deafult		: BOOL;
	st_SyncAuto		:BOOL	:=TRUE;		(* Piston state synchronized to last auto cycle command	*)
	set_SyncAuto	:BOOL;	
	b_Print_NotSyncAutoMessage :BOOL;
	
	//additional status for Upper and Lower
	st_Upper		:	BOOL	;
	st_Lower		:	BOOL	;

	// Each piston has its ID number
	iPisNum			:INT;
	
	DefaultCmd		:REFERENCE TO E_PistonDefault_CMD;

	// Timing 
	t_minOpen		:REFERENCE TO REAL;	(*Second*)	(* minimum time to open piston*)
	t_minClose		:REFERENCE TO REAL;	(*Second*)	(* minimum time to close piston*)
	t_maxOpen		:REFERENCE TO REAL;	(*Second*)	(* Maximum time to open piston, will initiate an error*)
	t_maxClose		:REFERENCE TO REAL;	(*Second*)	(* Maximum time to open piston, will initiate an error*)
	t_DelayOpen		:REFERENCE TO REAL;	(*Second*)	(* Delay time to getting "st_Open", will count after minimum time and sensors detection done*)
	t_DelayClose	:REFERENCE TO REAL;	(*Second*)	(* Delay time to getting "st_Close", will count after minimum time and sensors detection done*)	

	t_LastOpen		:TIME;			(* The last piston opening operation time*)
	t_LastClose		:TIME;			(* The last piston closing operation time*)
	
	//
	eErrNum			:E_ErrorPiton;		(* Error number*)
	sName			:STRING;		(* Piston description*)	
	
	//FB_Piston reference
	sen_Open: 		REFERENCE TO BOOL;
	sen_Close: 		REFERENCE TO BOOL;
	sen_Open_Exist: REFERENCE TO BOOL;
	sen_Close_Exist:REFERENCE TO BOOL;		
	
	valve_Open:		REFERENCE TO BOOL;
	valve_Close:	REFERENCE TO BOOL;	
	
	eModeZone:E_ModeZone;
END_STRUCT
END_TYPE

// ---- 00 Library/01 Piston/ST_Piston_SelectionList.TcDUT
TYPE ST_Piston_SelectionList :
STRUCT
	Num: INT;
	Description: STRING(80);

END_STRUCT
END_TYPE

// ---- 00 Library/01 Piston/ST_Piston_Setting_Param.TcDUT
TYPE ST_Piston_Setting_Param :
STRUCT

	// Timing 
	t_minOpen		:REAL 	:=1.5;	(*Second*)	(* minimum time to open piston*)
	t_minClose		:REAL	:=1.5;	(*Second*)	(* minimum time to close piston*)
	t_maxOpen		:REAL 	:=3.0;	(*Second*)	(* Maximum time to open piston, will initiate an error*)
	t_maxClose		:REAL	:=3.0;	(*Second*)	(* Maximum time to open piston, will initiate an error*)
	t_DelayOpen		:REAL 	:=0.0;	(*Second*)	(* Delay time to getting "st_Open", will count after minimum time and sensors detection done*)
	t_DelayClose	:REAL	:=0.0;	(*Second*)	(* Delay time to getting "st_Close", will count after minimum time and sensors detection done*)	

	sen_Open_Exist	: BOOL;
	sen_Close_Exist	: BOOL;		

END_STRUCT
END_TYPE

// ---- 00 Library/01 Piston/ST_Piston_U_L.TcDUT
TYPE ST_Piston_U_L :
STRUCT
	exist		: 	BOOL	; // true if device exist
	bError		:	BOOL	;
	iFB_Num		: E_Pis_Name;//Parent valve ID number

	//request
	req_Open	:	BOOL	;
	req_Close	:	BOOL	;
	req_Upper	:	BOOL	;
	req_Lower	:	BOOL	;
	req_None		:	BOOL	;
	
	//status
	st_Upper		:	BOOL	;
	st_Lower		:	BOOL	;
	st_Released		:	BOOL	;
	
	
	//Output
	out_Lower	:	BOOL	;
	out_Upper	:	BOOL	;
	
	//sensors
	sen_Upper			:	BOOL	;
	sen_Lower			:	BOOL	;	
	sen_Upper_exist		:	BOOL	;
	sen_Lower_exist		:	BOOL	;	
	//getting the structure of piston
	//str_Piston	:	REFERENCE TO ST_Piston	;
END_STRUCT
END_TYPE

// ---- 00 Library/02 Pump/ControlWordStruct.TcDUT
TYPE ControlWordStruct :
STRUCT
    SwitchOn           : BOOL;  // Bit 0: Switch on
    EnableVoltage      : BOOL;  // Bit 1: Enable voltage
    QuickStop          : BOOL;  // Bit 2: Quick stop
    EnableOperation    : BOOL;  // Bit 3: Enable operation
    Reserved1          : BOOL;  // Bit 4: Reserved
    Reserved2          : BOOL;  // Bit 5: Reserved
    Reserved3          : BOOL;  // Bit 6: Reserved
    Reserved4          : BOOL;  // Bit 7: Reserved
    FaultReset         : BOOL;  // Bit 8: Fault reset
    Reserved5          : BOOL;  // Bit 9: Reserved
    Reserved6          : BOOL;  // Bit 10: Reserved
    Reserved7          : BOOL;  // Bit 11: Reserved
    Reserved8          : BOOL;  // Bit 12: Reserved
    Reserved9          : BOOL;  // Bit 13: Reserved
    Reserved10         : BOOL;  // Bit 14: Reserved
    Reserved11         : BOOL;  // Bit 15: Reserved	
END_STRUCT
END_TYPE

// ---- 00 Library/02 Pump/StatusWordStruct.TcDUT
TYPE StatusWordStruct :
STRUCT
    ReadyToSwitchOn       : BOOL;  // Bit 0
    SwitchedOn            : BOOL;  // Bit 1
    OperationEnabled      : BOOL;  // Bit 2
    Fault                 : BOOL;  // Bit 3
    VoltageEnabled        : BOOL;  // Bit 4
    QuickStop             : BOOL;  // Bit 5
    SwitchOnDisabled      : BOOL;  // Bit 6
    Warning               : BOOL;  // Bit 7
    Remote                : BOOL;  // Bit 8
    Reserved1             : BOOL;  // Bit 9
    Reserved2             : BOOL;  // Bit 10
    Reserved3             : BOOL;  // Bit 11
    Reserved4             : BOOL;  // Bit 12
    Reserved5             : BOOL;  // Bit 13
    Reserved6             : BOOL;  // Bit 14
    Reserved7             : BOOL;  // Bit 15	
END_STRUCT
END_TYPE

// ---- 00 Library/02 Pump/ST_Pump.TcDUT
TYPE ST_Pump :
STRUCT
	//request
	modeAuto	:	BOOL	;//System in automatic
	bRun_Auto	:	BOOL	;
	bRun_Man	:	BOOL	;
	bRun		: 	BOOL;
	DriveReady	: 	BOOL;

	nRPM_Auto	:	REAL		;//Pump RPM 
	nRPM_Man	:	REAL		;//Pump RPM 
	nRPM		:	REAL		;//Pump RPM 
	//feedback
	nRPM_fdbk	:	INT	;
END_STRUCT
END_TYPE

// ---- 00 Library/03 SFC/ST_SFC.TcDUT
TYPE ST_SFC :
STRUCT
	SFCInit:		REFERENCE TO BOOL;
	SFCReset:		REFERENCE TO BOOL;
	SFCError:		REFERENCE TO BOOL;
	SFCEnableLimit:	REFERENCE TO BOOL;
	SFCErrorStep:	REFERENCE TO STRING;
	SFCErrorPOU:	REFERENCE TO STRING;
	SFCQuitError:	REFERENCE TO BOOL;
	SFCPause:		REFERENCE TO BOOL;
	SFCTrans:		REFERENCE TO BOOL;
	SFCCurrentStep:	REFERENCE TO STRING;
	SFCTip:			REFERENCE TO BOOL;
	SFCTipMode:		REFERENCE TO BOOL;
END_STRUCT
END_TYPE

// ---- 00 Library/04 Recipe/E_Recipe_Root_Folder.TcDUT
{attribute 'qualified_only'}
{attribute 'strict'}
TYPE E_Recipe_Root_Folder :
(
	PLC := 0,
	Develop_1,
	Develop_2,
	Develop_3,
	Develop_4	
);
END_TYPE

// ---- 00 Library/04 Recipe/ST_Recipe.TcDUT
TYPE ST_Recipe :
STRUCT
	arrRecipeNames 			:ARRAY[0..GVL_Recipe.C_Max_RecipeFileNum] OF STRING;//(20);
	arrVariableNamesValue 	:ARRAY[0..1200] OF STRING;//(40);
	arrVariableValue 		:ARRAY[0..1200] OF STRING;//(40);
	arrVariableDisp 		:ARRAY[0..2,0..20] OF STRING;//(40);


	sSelectedReceipe		:STRING(30);
	sLastSelectedReceipe	:STRING(30);
	sNewRecipeName			:STRING(30);
	//sRecipeDef				:STRING := 'Recipe'; (* current recipe definition *)
	iRecipeIndex 			:INT;
	iRecipeCount			:INT;
	bSaveFileCmd			:BOOL;
	bWriteToPLC_Cmd			:BOOL;
	bValidSelected			:BOOL;
	bCreateRecipe			:BOOL;
	bDeleteRecipe			:BOOL;
	bReloadRecipes			:BOOL:=TRUE;
	bInit					:BOOL:=FALSE;;
	bReInit					:BOOL;
	bShowFile				:BOOL;
	bGetLastError			:BOOL;
	bResetLastError			:BOOL;
	iDispSel				:INT; // 0..1180 --- 1200-20=1180 - Scrollbar fot HMI Table name & value
	info					:InfoValues;
	
END_STRUCT
END_TYPE

// ---- 00 Library/04-Messages/DUTs/Errors/E_ErrorFormat.TcDUT
TYPE E_ErrorFormat :(
	eErrID:=0,
	eErrLevel:=1,
	eErrMeassage:=2,
	eErrModuleDescription:=3
);
END_TYPE

// ---- 00 Library/04-Messages/DUTs/Errors/ST_Error.TcDUT
TYPE ST_Error :
STRUCT
	b_Active				: BOOL;
	b_memo				: BOOL;
	(*e_Description			: E_ErrorList;*)
	iErNum				: INT;
END_STRUCT
END_TYPE

// ---- 00 Library/04-Messages/DUTs/Errors/ST_Mess_Logger.TcDUT
TYPE ST_Mess_Logger :
STRUCT
	iErNum					: INT;
	sTime					: STRING[20];
	sDate					: STRING[20];
	sDescription				: STRING[40];
END_STRUCT
END_TYPE

// ---- 00 Library/04-Messages/DUTs/stMessageFormat.TcDUT
TYPE stMessageFormat :
STRUCT
	sDateTime							: STRING[25];
	sErrID								: STRING[11];
	sLevel								: STRING[10];
	sModuleDescription					: STRING[80];
	sErrorMessage						: STRING[200];	
END_STRUCT
END_TYPE

// ---- 00 Library/05 Safety/ST_ES_PB.TcDUT
TYPE ST_ES_PB :
STRUCT
	in: BOOL;
	State: BOOL;
	Memo: BOOL;
	ByPass: BOOL;
	stBitMap                : STRING:= 'ImagePool.EStop_OK2'; //'ImagePool.EStop_ACT2'
END_STRUCT
END_TYPE

// ---- 00 Library/05 Safety/ST_SafeOut_PlcIn.TcDUT
TYPE ST_SafeOut_PlcIn :
STRUCT
	ES1_PB_State	:BOOL;
	ES2_PB_State	:BOOL;
	ES3_PB1_State	:BOOL;
	ES3_PB2_State	:BOOL;
	ES4_PB_State	:BOOL;
	
	ES1_State		: BOOL;
	ES2_State		: BOOL;
	ES3_State		: BOOL;
	ES4_State		: BOOL;
	
	TankLocked_CIP_T91: BOOL;
	TankLocked_CIP_T92: BOOL;
	TankLocked_CIP_T93: BOOL;
	TankLocked_CIP_T94: BOOL;
	TankLocked_Marinade_T1: BOOL;
	TankLocked_Marinade_T2: BOOL;
	TankLocked_Color_T3: BOOL;
	TankLocked_Color_T4: BOOL;

END_STRUCT
END_TYPE

// ---- 00 Library/05 Safety/ST_SafeIn_PlcOut.TcDUT
TYPE ST_SafeIn_PlcOut :
STRUCT
	ES1_PB_Restart						:BOOL;
	ES2_PB_Restart						:BOOL;
	ES3_PB_Restart						:BOOL;
	ES4_PB_Restart						:BOOL;
	
	ES1_HMI_PB_Button						:BOOL:=TRUE;
	ES2_HMI_PB_Button						:BOOL:=TRUE;
	ES3_HMI_PB_Button						:BOOL:=TRUE;
	ES4_HMI_PB_Button						:BOOL:=TRUE;
	
END_STRUCT
END_TYPE

// ---- 00 Library/05 Safety/TwinSAFE/e_DualChanal.TcDUT
TYPE e_DualChanal :(
	Wrong:=0,
	Close:=1,
	Open:=2);
END_TYPE

// ---- 00 Library/05 Safety/TwinSAFE/TwinSafeOut_PlcIn.TcDUT
TYPE TwinSafeOut_PlcIn :
STRUCT
	FB_Err			: BOOL;
	COM_Err			: BOOL;
	OUT_Err			: BOOL;
	Other_Err		: BOOL;
	InRun			: BOOL;
	//ES_State		: BOOL;

END_STRUCT
END_TYPE

// ---- 00 Library/05 Safety/TwinSAFE/TwinSafeIn_PlcOut.TcDUT
TYPE TwinSafeIn_PlcOut :
STRUCT
	RUN			: BOOL;
	ErrACK		: BOOL;
	//Restart		: BOOL; //Restart TwinSAFE
END_STRUCT
END_TYPE

// ---- 00 Library/07 Errors/E_Error_Active_Module.TcDUT
{attribute 'qualified_only'}
{attribute 'strict'}
TYPE E_Error_Active_Module :
(
	noError := 0, Piston, Motor
);
END_TYPE

// ---- 00 Library/07 Errors/E_OwnerDevice.TcDUT
{attribute 'qualified_only'}
{attribute 'strict'}
TYPE E_OwnerDevice :
(
	NotDefined := 0,
	Tank1,
	Tank2,
	Tank3,
	Tank4,
	common //last
);
END_TYPE

// ---- 00 Library/07 Errors/ST_DeviceErrorHandeling.TcDUT
TYPE ST_DeviceErrorHandeling :
STRUCT
	eName			: E_OwnerDevice:=E_OwnerDevice.NotDefined;
	sObjectName		: STRING:='Device Name';
	iObjectID		: INT;
	sLastErrorStep	: STRING;
	eErrorActive	: E_Error_Active_Module:=E_Error_Active_Module.noError;
	bMasterResume	: BOOL;

END_STRUCT
END_TYPE

// ---- 00 Library/07-Mode/E_BuzzerMode.TcDUT
TYPE E_BuzzerMode :
(
	eBuzzerOff := 0,
	eBuzzerError,		//Short Delay Off
	eBuzzerWarning		//Long Delay Off
);
END_TYPE

// ---- 00 Library/07-Mode/E_LightTowerState.TcDUT
TYPE E_LightTowerState :
(
	eLightsOff:=0,
	eGreen,						//Run All
	eGreen_YellowBlink,			//Run All and warning
	eGreenBlink,				//Run some and some not
	eGreenBlink_YellowBlink,	//Run some and warning
	eGreenBlink_RedBlink,		//Run some and error
	eYellow,					//Pause
	eBlue,						//
	eRed						//Error
);
END_TYPE

// ---- 00 Library/07-Mode/E_OperationButtons.TcDUT
TYPE E_OperationButtons :(
	ePauseAll:=0,
	ePlayAll:=1);
END_TYPE

// ---- 00 Library/07-Mode/E_WorkingMode.TcDUT
TYPE E_WorkingMode :(	
	eManualMode			:=0,
	eSemiAutoMode		:=1,
	eAutoMode			:=2);
END_TYPE

//eWorkingModeNone	:=0,

// ---- 00 Library/07-Mode/ST_Mode.TcDUT
TYPE ST_Mode :
STRUCT
	iActMode: E_WorkingMode;
	bSetManual: BOOL;
	bSetSemi: BOOL;
	bSetAuto: BOOL;

	eModeZone:E_ModeZone:=E_ModeZone.eNone;
	
	bStateSafe_mode: BOOL:=TRUE;

END_STRUCT
END_TYPE

// ---- 00 Library/07-Mode/ST_OperationButtons.TcDUT
TYPE ST_OperationButtons :
STRUCT
	iActOperation	: E_OperationButtons;
	bSetPause		: BOOL;
	bSetPlay		: BOOL;
	bResetError		: BOOL;
	bStopResetAll	: BOOL;
	bPauseOnDelayed	: BOOL;
	
	bStateSafe_mode : BOOL:=TRUE;
	
	b_rt_Pause		: BOOL;
	b_rt_Play		: BOOL;	

	eModeZone		: E_ModeZone;
	sModeZone		: STRING;
	iPauseHistory	: INT;
	
	iActModeState	: E_WorkingMode; //just for reference stete not for change 
END_STRUCT
END_TYPE

// ---- 00 Library/11 HMI/E_Led_Color.TcDUT
{attribute 'qualified_only'}
{attribute 'strict'}
{attribute 'to_string'}
TYPE E_Led_Color :
(
	Yellow := 0,
	Red,
	Green,
	Blue,
	Gray
	
);
END_TYPE

// ---- 00 Library/11 HMI/ST_MixProof_state.TcDUT
TYPE ST_MixProof_state :
STRUCT
	sName: STRING;
	bUpper: BOOL;
	bLower: BOOL;
	bRunning: BOOL;
	bDone: BOOL;

END_STRUCT
END_TYPE

// ---- 00 Library/12 Analog Sensor/E_ASensor_State.TcTLEO
{attribute 'qualified_only'}
{attribute 'strict'}
TYPE E_ASensor_State :
(
	Init := 0,
	Close,Open,Busy_Close,Busy_Open
);
END_TYPE

// ---- 00 Library/12 Analog Sensor/ST_AnalogSensor.TcDUT
TYPE ST_AnalogSensor :
STRUCT
	ID		: STRING;
	Value	: REAL;
	Unit	: STRING;
	
	//rawVal_Sensor	: REAL;
	rawVal_Min		: REAL;
	rawVal_Max		: REAL;
	
	outVal_Min		: REAL;
	outVal_Max		: REAL;
	outOffset		: REAL;
	
	//alarms warning
	rLL_Alarm		: REAL	;
	rHH_Alarm		: REAL	;
	rLL_Warning		: REAL	;
	rHH_Warning		: REAL	;
	
END_STRUCT
END_TYPE

// ---- 00 Library/13 Process Control/ST_ProcessControl.TcDUT
TYPE ST_ProcessControl :
STRUCT
	idName			: STRING;

	rValue			: REAL;
	rSetPoint		: REAL;
	Deviation		: REAL;
	rValue_Min_To_ReleaseControl		: REAL;
	
	ToleravceLow	: REAL:=0;  // min=0
	ToleranceHigh	: REAL:=0;  // min=0

	Control_Value	: REAL;  // min=0 , max=1
	Control_ON		: BOOL;
	OverFlow		: BOOL;	
	
	//PID parameters
	bPause			: 	BOOL	;
	bManual			: 	BOOL	;
	bReset			: 	BOOL	;
	fCtrlCycleTime	: 	REAL	; 
	fKp				:	REAL	; 
	fTn				:	REAL	; 
	fTv				:	REAL	;
	fTd				:	REAL	; // not in use
	fCtrlOutput		:	LREAL	; 
	fCtrlOutput_Manual		:	LREAL	; 
	fCtrlOutput_Min			:	LREAL:=300	; 
	fCtrlOutput_Max			:	LREAL:=3000	; 

	nErrorStatus 	: 	UINT	;
	
	//Hysteresis
	fHystHigh		:	REAL	;
	fHystLow		:	REAL	;
	bHystOut		:	BOOL	;
	rHystOutLow		:	REAL:=1200	;
	rHystOutHigh	:	REAL:=2500	;
	
	bDone			:	BOOL	;
	bActiveCntr		:	BOOL	;
	
	nNumberOfDcNum	:	INT	;//Number of number after decimal point
END_STRUCT
END_TYPE

// ---- 00 Library/30 IO/ST_EL3xx8.TcDUT
TYPE ST_EL3xx8 :
STRUCT
	ch1		:INT;
	ch2		:INT;
	ch3		:INT;
	ch4		:INT;
	ch5		:INT;
	ch6		:INT;
	ch7		:INT;
	ch8		:INT;
END_STRUCT
END_TYPE

// ---- 00 Library/30 IO/ST_EL18x9.TcDUT
TYPE ST_EL18x9 :
STRUCT
	
	State	AT %I*: UINT;
	i_ch1	AT %I*: BOOL;
	i_ch2	AT %I*: BOOL;
	i_ch3	AT %I*: BOOL;
	i_ch4	AT %I*: BOOL;
	i_ch5	AT %I*: BOOL;
	i_ch6	AT %I*: BOOL;
	i_ch7	AT %I*: BOOL;
	i_ch8	AT %I*: BOOL;
	
	i_ch9	AT %I*: BOOL;
	i_ch10	AT %I*: BOOL;
	i_ch11	AT %I*: BOOL;
	i_ch12	AT %I*: BOOL;
	i_ch13	AT %I*: BOOL;
	i_ch14	AT %I*: BOOL;
	i_ch15	AT %I*: BOOL;
	i_ch16	AT %I*: BOOL;
	
END_STRUCT
END_TYPE

// ---- 00 Library/30 IO/ST_EL1918_TwinSafe.TcDUT
TYPE ST_EL1918_TwinSafe :
STRUCT
	
//EtherCAT Terminal, 8-channel digital input, 
//24 V DC, TwinSAFE, TwinSAFE Logic

	State	AT %I*: UINT;
	i_ch1	AT %I*: BOOL;
	i_ch2	AT %I*: BOOL;
	i_ch3	AT %I*: BOOL;
	i_ch4	AT %I*: BOOL;
	i_ch5	AT %I*: BOOL;
	i_ch6	AT %I*: BOOL;
	i_ch7	AT %I*: BOOL;
	i_ch8	AT %I*: BOOL;
	
END_STRUCT
END_TYPE

// ---- 00 Library/30 IO/ST_EL28x9.TcDUT
TYPE ST_EL28x9 :
STRUCT
	//16CH DO, PNP 24VDC/0.5A  - 2809
	//16CH DO, GND-SW, 24VDC/0.5A - 2889
	
	State	AT %I*: UINT;

	q_ch1	AT %Q*: BOOL;
	q_ch2	AT %Q*: BOOL;
	q_ch3	AT %Q*: BOOL;
	q_ch4	AT %Q*: BOOL;
	q_ch5	AT %Q*: BOOL;
	q_ch6	AT %Q*: BOOL;
	q_ch7	AT %Q*: BOOL;
	q_ch8	AT %Q*: BOOL;
	
	q_ch9	AT %Q*: BOOL;
	q_ch10	AT %Q*: BOOL;
	q_ch11	AT %Q*: BOOL;
	q_ch12	AT %Q*: BOOL;
	q_ch13	AT %Q*: BOOL;
	q_ch14	AT %Q*: BOOL;
	q_ch15	AT %Q*: BOOL;
	q_ch16	AT %Q*: BOOL;
	
(*	
	bit_ch1	AT %Q*: BIT;
	bit_ch2	AT %Q*: BIT;
	bit_ch3	AT %Q*: BIT;
	bit_ch4	AT %Q*: BIT;
	bit_ch5	AT %Q*: BIT;
	bit_ch6	AT %Q*: BIT;
	bit_ch7	AT %Q*: BIT;
	bit_ch8	AT %Q*: BIT;
	
	bit_ch9		AT %Q*: BIT;
	bit_ch10	AT %Q*: BIT;
	bit_ch11	AT %Q*: BIT;
	bit_ch12	AT %Q*: BIT;
	bit_ch13	AT %Q*: BIT;
	bit_ch14	AT %Q*: BIT;
	bit_ch15	AT %Q*: BIT;
	bit_ch16	AT %Q*: BIT;
*)	
	
	
	
END_STRUCT
END_TYPE

// ---- 00 Library/30 IO/ST_EL2904.TcDUT
TYPE ST_EL2904 :
STRUCT
	State	AT %I*: UINT;
	q_ch1	AT %Q*: BOOL;
	q_ch2	AT %Q*: BOOL;
	q_ch3	AT %Q*: BOOL;
	q_ch4	AT %Q*: BOOL;
	
END_STRUCT
END_TYPE

// ---- 00 Library/30 IO/ST_EL3xx4.TcDUT
TYPE ST_EL3xx4 :
STRUCT
	
	//4CH AI, RTD RES SNS
	State	AT %I*: UINT;

	ai_ch1	AT %I*: INT;
	ai_ch2	AT %I*: INT;
	ai_ch3	AT %I*: INT;
	ai_ch4	AT %I*: INT;
	
	
END_STRUCT
END_TYPE

// ---- 00 Library/30 IO/ST_EL4xx8.TcDUT
TYPE ST_EL4xx8 :
STRUCT
	ch1		:INT;
	ch2		:INT;
	ch3		:INT;
	ch4		:INT;
	ch5		:INT;
	ch6		:INT;
	ch7		:INT;
	ch8		:INT;
END_STRUCT
END_TYPE

// ---- 00 Library/30 IO/ST_Nidec.TcDUT
TYPE ST_Nidec :
STRUCT
	StatusWord     AT %I* : WORD;     // Input from Receive PDO Mapping 6
	ControlWord     AT %Q* : WORD;      // Output to Transmit PDO Mapping 6
	
	actVelocity AT %I*: INT;
	targetVelocity AT %Q*: INT;
END_STRUCT
END_TYPE

// ---- 00 Library/30 IO/ST_TwinSAFE.TcDUT
TYPE ST_TwinSAFE :
STRUCT
	TSafeIn			AT %I*	: TwinSafeOut_PlcIn;
	TSafeOut		AT %Q*	: TwinSafeIn_PlcOut;
	stSafetyIn		AT %I* 	: ST_SafeOut_PlcIn;
	stSafetyOut		AT %Q* 	: ST_SafeIn_PlcOut;	
END_STRUCT
END_TYPE

// ---- 00 Library/30 IO/ST_VTUG.TcDUT
TYPE ST_VTUG :
STRUCT
	sol_14: BOOL;
	sol_12: BOOL;
END_STRUCT
END_TYPE

// ---- 00 Library/HeatExchenger/ST_HeatExchanger.TcDUT
TYPE ST_HeatExchanger :
STRUCT
	//request
	bManual	:	BOOL	;//System in automatic
	bRun	:	BOOL	;
	nTemp	:	INT		;
	//feedback
	nTemp_fdbk	:	INT	;
	
	//Output signal scaling
	cntrlVal_Min		: REAL:=0;
	cntrlVal_Max		: REAL:=100;
	
	outVal_Min		: REAL:=0;
	outVal_Max		: REAL:=32767;
	outOffset		: REAL:=0;
	fManualControl	: LREAL:=100;

END_STRUCT
END_TYPE

// ---- 00 Library/Sensors/E_Tank_Level.TcDUT
{attribute 'qualified_only'}
{attribute 'strict'}
TYPE E_Tank_Level :
(
	eEmpty := 0,
	eLL,
	eHL,
	eERROR
	
);
END_TYPE

// ---- 00 Library/Sensors/ST_AnalogSignal.TcDUT
TYPE ST_AnalogSignal :
STRUCT
	//analog signal
	nIn_RawSignal	:	UINT		;
	rOut_Converted	:	REAL	;
	
	//analog signal settings
	rRawMax	:	REAL:=32767	;
	rRawMin	:	REAL:=0		;
	rOutMax	:	REAL:=100	;
	rOutMin	:	REAL:=10 	;
	//not usable 
	rRawZeroPointOffset	:	REAL:=100;//offset foranalog signal //?
	rRawMaxPointOffset	:	INT:=100;//?
END_STRUCT
END_TYPE

// ---- 00 Library/Sensors/ST_Tank_Level.TcDUT
TYPE ST_Tank_Level :
STRUCT
	//Input signals fro I/O
	bIn_LL_signal	:	BOOL :=TRUE	;
	bIn_HL_signal	:	BOOL :=TRUE	;
	//Tank level state, empty, Low level, High level
	e_state			:	E_Tank_Level:=E_Tank_Level.eHL	;
	
	rTankLevel				:	REAL	;
	rTankLevelPercentage	:	REAL	;
END_STRUCT
END_TYPE

// ---- 01 Instance/01 Piston/E_Pis_Name.TcDUT
{attribute 'qualified_only'}
//{attribute 'strict'}
{attribute 'to_string'}
TYPE E_Pis_Name :
(
	e0_not_in_use := 0,
	// CIP Source
	V1001,
	V1002,
	V1003,
	V1004,
	V1005,

	MV1001,
	MV1002,
	MV1003,
	MV1004,
	
	//CIP Return
	V1101,
	V1102,
	V1103,
	V1104,
	V1105,
	V1112,
	V1114,
	V1117,
	V1120,
	
	//CIP Client
	V1106,
	V1023,V1024,V1025,V1026,V1027,V1028,V1029,V1030,

	//CIP Client Tanks
	V3001,V3003,V3005,V3006,V3007,V3041,V3039,
	V4001,V4003,V4005,V4006,V4007,V4041,V4039,	
	
	//CIP Tanks
	V1011,V1012,V1013,
	V1014,V1015,V1016,
	V1017,V1018,V1019,
	V1020,V1021,V1022,
	V1031,V1032,
	
	//Tank Target 1
	V3016,
	V3017,
	V3023,
	V3024,
	V3025,
	V3026,	
	
	//Tank Target 2
	V3015,	
	V3027,	
	V3028,	
	V3029,	
	V3030,	
	
	//Marinade Lines
	V3018,
	V3019,
	V3020,V3040,
	V3021,
	V3022,
	
	V3014,
	V3113,
	
	
	
	//Tank Target 3
	V4016,
	V4017,
	V4023,
	V4024,
	V4025,
	
	//Tank Target 4
	V4015,
	V4026,
	V4027,
	V4028,
	V4029,
	V4030,
	
	//Color Lines
	V4018,
	V4019,
	V4020,V4040,
	V4021,
	V4022,
	
	V2115,
	V2116,
	V2117,
	
	// Tanks Coolant
	V3031,V3032,
	V3033,V3034,
	V4031,V4032,
	V4042,V4043,
	
	//TriBlender Select
	V3035,V4037,V5001,
	V3038,V4038,V5002,
	
	//addition
	
	V4014,
	V4113,
	V2114,
	
	V3004,
	V3008,
	V3009,
	V3010,
	
	V4034,
	V4033,
	V4035,
	V4036,
	
	V4004,
	V4010,
	V4008,
	V4009,
	
	//Water
	V2011,V2111,V2211,V2112,
	
	
	V5012,
	
	V4026_2, //temp for marinade filling test 
	
	//Dummy valves for fbLineTarget_Marinade
	V_Dummy_01,
	V_Dummy_02,
	V_Dummy_03,
	V_Dummy_04,
	V_Dummy_05,
	V_Dummy_06,
	V_Dummy_07,
	V_Dummy_08,
	V_Dummy_09,
	V_Dummy_10,
	V_Dummy_11,
	V_Dummy_12,
	
	//Dummy for Line Source Marinada
	V_Dummy_LSM_01,
	V_Dummy_LSM_02,
	V_Dummy_LSM_03,
	V_Dummy_LSM_04,
	V_Dummy_LSM_05,
	V_Dummy_LSM_06,
	V_Dummy_LSM_07, //*
	//Dummy for TriBlender Source Marinada
	V_Dummy_TSM_01,
	V_Dummy_TSM_02,
	V_Dummy_TSM_03,
	//Dummy for Line Source Color
	V_Dummy_LSC_01,
	V_Dummy_LSC_02,
	V_Dummy_LSC_03,
	V_Dummy_LSC_04, //*
	
	//Dummy Drain Tap Water
	V_Dummy_DTW_01,
	
	
	//virtual list
	last
	



	
);
END_TYPE

// ---- 01 Instance/02 Pump/E_Pump_List.TcDUT
{attribute 'qualified_only'}
{attribute 'strict'}
{attribute 'to_string'}
TYPE E_Pump_List :
(
	eNotSelected := 0,
	P1001,
	P3001,
	P3002,
	P4001, //Line Color
	P4002, //CIP Color return
	TB0001,
	PP1002,
	PP1003,
	AG3001,
	AG3002,
	AG4001,
	AG4002,
	
	
	last
);
END_TYPE

// ---- 01 Instance/04 Recipe/E_Recipe_Name.TcDUT
//{attribute 'qualified_only'}
//{attribute 'strict'}
{attribute 'to_string'}
TYPE E_Recipe_Name :
(
	//e0_not_in_use := 0,
	R_All:=1,
	R_Device_Dough1,
	R_Device_Dough2,
	R_Device_Dough3,
	R_Device_Dough4,
	R_Piston_Settings // must be last
	
);
END_TYPE

// ---- 01 Instance/07-Mode/E_LightTower_Type.TcDUT
{attribute 'qualified_only'}
{attribute 'strict'}
TYPE E_LightTower_Type :
(
	eSingleLayer := 0,
	eMultiLayer
);
END_TYPE

// ---- 01 Instance/07-Mode/E_ModeZone.TcDUT
{attribute 'qualified_only'}
{attribute 'strict'}
{attribute 'to_string'}
TYPE E_ModeZone :
(
	eNone := 0,
	eMain,
	
	eCIP,
	eTank1,(*Tank*)
	eTank2,(*Tank*)
	eTank3,(*Tank*)
	eTank4,(*Tank*)
	
	eProduction_Marinade,(*Line*)
	eProduction_Color,(*Line*)
	
	eTriBlender_Marinade,(*Line*)
	eTriBlender_Color,(*Line*)
	eWater,(*Line*)
	eHotWater,(*Line*)
	eLast
);
END_TYPE

// ---- 01 Instance/07-Mode/E_SkidZone.TcDUT
{attribute 'qualified_only'}
{attribute 'strict'}
TYPE E_SkidZone :
(
	eCIP := 0,
	eTriBlender,
	eMarinade,
	eColor,
	eLast
);
END_TYPE

// ---- 01 Instance/12 Analog Sensor/E_ASense_Name.TcTLEO
{attribute 'qualified_only'}
{attribute 'strict'}
{attribute 'to_string'}
TYPE E_ASense_Name :
(
	eNotSelected := 0,
	//level sensors CIP	
	LT1004,	
	LT1003,	
	LT1002,
	LT1001,
	//Flow  sensors
	FT1001,
	FT1002,

	
	
	//conductivity sensors
	CT1101,
	CT3101,//not exist	
		
	//temperature sensors
	TT1001,
	TT1002,
	TT1003,
	TT1004,
	TT1101,
	TT1105,
	CT1101_2,
	CT1101_3,
	CT1101_4,
	TT2001,
	TT3001,
	TT3002,
	TT4001,
	TT4002,
	
	//level sensors


	LT1061,
	LT1071,
	LT3001,
	LT3002,
	LT4001,
	LT4002,
	
	//Pressure sensors
	PT1001,
	PT3001,
	PT3002,
	PT4001,
	PT4002,
	PT9001,
	PT9002,
	PT9011,

	FT4001,
	FT4002,	
	FT9011,
	
	//Air Pressure
	AP1001, //CIP
	AP2001, // TriBlender
	AP3001, //Marinade
	AP4001, //Color
	
	CT4101,	
	CT4102,	

	FT9012,
	
	//virtual list
	last
);
END_TYPE

// ---- 01 Instance/13 Process Control/E_ProcessControl_Name.TcDUT
{attribute 'qualified_only'}
{attribute 'strict'}
{attribute 'to_string'}
TYPE E_ProcessControl_Name :
(
	(*
	888888
	888888 NOTE !!! add new element ONLY before the last element <eProcCntrl_Last>!!!
	888888
	*)
	e0_not_in_use := 0,
	//Concentration
	eDetergentConc,		//Detergent concentration
	eDisinfectionConc,	//Disinfection concentration
	//Temperature
	eDeterTemp, //Detergent temperature
	eDisTemp,	//Disinfection temperature
	eMarinTank1_Temp,
	eMarinTank2_Temp,
	eColorTank1_Temp,
	eColorTank2_Temp,
	eClientReturn_Temp,
	//Flow rate
	eCIP_Flow_1,//**FT1001 CIP
	eCIP_Flow_2,//**FT1002 CIP Client return pipe
	eCIP_Flow_3,//**FT1002 CIP Client return sprinkler
	
	//Level
	eMarin_Level,
	eColor_Level,
	//Pressure
	eCIP_Pressure,
	
	eHeatExchanger,
(*	
	eTriBlender_Flow,//**FT9011
	
	eColor_TriB_Conc,//**CT4101
	eColor_Line_Conc,//**CT4102

	eP3001_Pressure,//**PT3001
	eP3002_Pressure,//**PT3002
	eP4001_Pressure,//**PT4001
	eP4002_Pressure,//**PT4002
*)	
	
	// add new element ONLY hire !!!
	eProcCntrl_Last
);
END_TYPE

// ---- 03 Project/23 CIP/E_Tank_Name.TcTLEO
{attribute 'qualified_only'}
{attribute 'strict'}
TYPE E_Tank_Name :
(
	enum_member := 0,
	
	//CIP
	T91,
	T92,
	T93,
	T94,
	
	//Marinade
	T1,
	T2,
	
	//Color
	T3,
	T4,
	
	last
	
);
END_TYPE

// ---- 03 Project/21 Data/E_Element_State_Long.TcDUT
{attribute 'qualified_only'}
//{attribute 'strict'}
{attribute 'to_string'}
TYPE E_Element_State_Long :
(
eOff := 0,
eStandby,
eNotClean,
eCIP_1_Rinzed,
eCIP_2_Deterged,
eCIP_3_Deterged_Clean,
eCIP_4_Sanitized,
eCIP_5_Done,
eWaterReady,
eReady,
eProduction,
// jump to eReady
eEmpty,
eExpired
);
END_TYPE

// ---- 03 Project/23 CIP/E_CIP_Client_Command.TcDUT
{attribute 'qualified_only'}
{attribute 'strict'}
TYPE E_CIP_Client_Command :
(
	eDrain := 0,
	eCIP,
	eClose
);
END_TYPE

// ---- 03 Project/23 CIP/E_CIP_Client_Selector.TcDUT
{attribute 'qualified_only'}
{attribute 'strict'}
TYPE E_CIP_Client_Selector :
(
	eNone := 0,
	eClose,
	eFuture,
	eMarinade_Up,
	eMarinade_Low,
	eColor_Up,
	eColor_Low,
	eDrain,
	eLoop
);
END_TYPE

// ---- 03 Project/23 CIP/E_CIP_DashStage.TcDUT
{attribute 'qualified_only'}
{attribute 'strict'}
TYPE E_CIP_DashStage :
(
	eCIPStage_NotInUse:= 0,
	eCIPStage_NotAvalable,
	eCIPStage_ToBeDone,
	eCIPStage_Active,
	eCIPStage_Done
);
END_TYPE

// ---- 03 Project/23 CIP/E_CIP_DashStage_List.TcDUT
{attribute 'qualified_only'}
//{attribute 'strict'}
{attribute 'to_string'}
TYPE E_CIP_DashStage_List :
(
	e00_NotSelected := 0,
	
	//CIP1
	e01_CIP1_Client_Drain_Product_Rest_Pipe,
	e02_CIP1_Client_Drain_Product_Rest_Sprinkler,
	
	//CIP2
	e03_CIP2_Local_Detergent_Fill,
	e04_CIP2_Local_Detergent_Condition,
	e05_CIP2_Client_Detergent_Fill,
	e06_CIP2_Client_Detergent_Condition_Pipe,	
	e07_CIP2_Client_Detergent_Condition_Sprinkler,	
	
	//CIP3
	e08_CIP3_Detergent_Collect,
	e09_CIP3_Detergent_Drain,
	e10_CIP3_Detergent_Clean_Pipe,
	e11_CIP3_Detergent_Clean_Sprinkler,
	
	//CIP4
	e12_CIP4_Local_DisInfection_Fill,
	e13_CIP4_Local_DisInfection_Condition,
	e14_CIP4_Client_DisInfection_Fill,
	e15_CIP4_Client_DisInfection_Condition_Pipe,	
	e16_CIP4_Client_DisInfection_Condition_Sprinkler,	
	
	//CIP5
	e17_CIP5_DisInfection_Collect,
	e18_CIP5_DisInfection_Drain,
	e19_CIP5_DisInfection_Clean_Pipe,
	e20_CIP5_DisInfection_Clean_Sprinkler,	
	
	
	eLast
);
END_TYPE

// ---- 03 Project/23 CIP/E_CIP_Mode.TcDUT
{attribute 'qualified_only'}
{attribute 'strict'}
TYPE E_CIP_Mode :
(
	eOff :=0,
	eManual,
	eAuto	
);
END_TYPE

// ---- 03 Project/23 CIP/E_CIP_Return.TcDUT
{attribute 'qualified_only'}
{attribute 'strict'}
TYPE E_CIP_Return :
(
	eNone := 0,
	eDrain,
	eT91_Sanitation,
	eT92_Detergent,
	eT93_R_Water,
	eT94_Water
);
END_TYPE

// ---- 03 Project/23 CIP/E_CIP_Source.TcDUT
{attribute 'qualified_only'}
{attribute 'strict'}
TYPE E_CIP_Source :
(
	eNone := 0,
	eT91_Sanitation,
	eT92_Detergent,
	eT93_R_Water,
	eT94_Water,
	eClose
);
END_TYPE

// ---- 03 Project/23 CIP/E_CIP_TankList.TcDUT
{attribute 'qualified_only'}
{attribute 'strict'}
TYPE E_CIP_TankList :
(
	eT91_Sanitation :=0,
	eT92_Detergent,
	eT93_R_Water,
	eT94_Water
);
END_TYPE

// ---- 03 Project/23 CIP/E_CIP_Type.TcDUT
{attribute 'qualified_only'}
{attribute 'strict'}
TYPE E_CIP_Type :
(
	NotSelected := 0,
	R_Water,
	Detergent,
	Full
);
END_TYPE

// ---- 03 Project/23 CIP/E_CIP_Usage.TcDUT
{attribute 'qualified_only'}
//{attribute 'strict'}
{attribute 'to_string'}
TYPE E_CIP_Usage :
(
	eNotInUse := 0,
	eTank_1,
	eTank_2,
	eTank_3,
	eTank_4,
	eTriBlender_Marinada,
	eTriBlender_Color,
	eLine_Marinada,
	eLine_Color,
	eLocal,
	eExternal	//GAD client through Siemens, stays after eLocal: arr_CIP_Param ends at eLocal
	//,eClient
);
END_TYPE

// ---- 03 Project/23 CIP/ST_CIP_Param.TcDUT
TYPE ST_CIP_Param :
STRUCT	//st_CIP_Param
	//New parameters
	sName: STRING;
	r_Tank91_Volume			:	REAL:=300	;	//volume in litres
	r_Tank92_Volume			:	REAL:=300	;	//volume in litres
	r_Tank93_Volume			:	REAL:=300	;	//volume in litres
	r_Tank94_Volume			:	REAL:=300	;	//volume in litres
	
	r_CIP_Pump				:	REAL:=200	;
	r_CIP_Client_Pump		:	REAL:=200	;
	
(**)r_Flow_Pipe				:	REAL:=160	;
(**)r_Flow_Sprinkler		:	REAL:=100	;
	
	r_Pressure				:	REAL:=0.5	;
	
	r_DetergentConcentration		:	REAL:=0.3	;//concentration in percents
	r_DisInfectionConcentration		:	REAL:=0.3	;//concentration in percents
	
	t_Measure_Delay						:	INT:=60		;//concentration measurment delay in seconds
(**)t_ConditionR_Water					:	INT:=60		;//concentration CIP time in seconds
(**)t_ConditionR_Water_Sprinkler		:	INT:=60		;//concentration CIP time in seconds
(**)t_ConditionDetergent				:	INT:=60		;//concentration CIP time in seconds
(**)t_ConditionDetergent_Sprinkler		:	INT:=60		;//concentration CIP time in seconds
(**)t_ConditionDisInfection				:	INT:=60		;//concentration CIP time in seconds
(**)t_ConditionDisInfection_Sprinkler	:	INT:=60		;//concentration CIP time in seconds
(**)t_ConditionWater					:	INT:=60		;//concentration CIP time in seconds
(**)t_ConditionWater_Sprinkler			:	INT:=60		;//concentration CIP time in seconds	
	r_Temper_Detergent					:	REAL:=65	;//temperature set point for local client in celsius
	r_Temper_DisInfection				:	REAL:=65	;//temperature set point for local client in celsius
(**)//r_Temper_ClientReturn				:	REAL:=65	;//Client return temperature
	t_PumpInitRun						:	INT:=20		;//pump initial run with constant RPM, time in seconds
(**)t_PumpInitRun_old					:	INT:=60		;(*not in use*)//pump start time in R_Water, time in seconds
	
(**)r_Volume_Sprinkler_Ratio		:	REAL:=0.7	;//in case of CIP Client Tanks, 0.7=70% of Volume to  sprinkler direction 
(**)r_Volume_Solution_Fill			:	REAL:=60	;//Client pipe volume displacement 
(**)r_Volume_Drain_R_Water			:	REAL:=20	;//Client pipe volume displacement 
	r_Volume_Collect_Detergent		:	REAL:=20	;//Client pipe volume displacement 
	r_Volume_Drain_Detergent		:	REAL:=20	;//Client pipe volume displacement 
	r_Volume_Recycle_Detergent		:	REAL:=20	;//Client pipe volume displacement 
	r_Volume_Collect_DisInfection	:	REAL:=20	;//Client pipe volume displacement 
	r_Volume_Drain_DisInfection		:	REAL:=20	;//Client pipe volume displacement 
	r_Volume_Recycle_DisInfection	:	REAL:=20	;//Client pipe volume displacement 

	(*//R_Water
		r_RWater_93_TankLvl	:	REAL:=150	;
		t_RWater_Pump_01	:	INT:=30		;//time in seconds
	
	//Detergent
		r_Deter_92_TankLvl_1	:	REAL:=250	;
		r_Deter_92_TankLvl_2	:	REAL:=300	;
		r_Deter_Flow_Pmp1_1		:	REAL:=200	;
		r_Deter_Flow_Pmp1_2		:	REAL:=200	;
		r_Deter_Pressure_Pmp1_1	:	REAL:=0.5	;
		n_Deter_PumpCIP_RPM		:	INT:=1500	;
		n_Deter_PumpClient_RPM	:	INT:=1500	;
		n_Deter_PumpCIP_RPM_1		:	INT:=1000	;
		n_Deter_PumpClient_RPM_1	:	INT:=1000	;
		
		//local
		st_Deter_Local			:	str_ConcParam	;
		//client
		st_Deter_Client			:	str_ConcParam	;
	
	//DisInfection
		r_DisInf_PumpCIP_RPM_1		:	INT:=1000	;
		r_DisInf_PumpCIP_RPM_2		:	INT:=1000	;
		r_DisInf_PumpClient_RPM_2	:	INT:=1000	;
		r_DisInf_PumpCIP_RPM_3		:	INT:=1000	;
		r_DisInf_PumpClient_RPM_3	:	INT:=1000	;
		//local
		st_DisInf_Local			:	str_ConcParam	;
		//client
		st_DisInf_Client		:	str_ConcParam	;
		
	//Water
		r_Water_TankLvl_Lcl_1		:	REAL:=250		;
		r_Water_TankLvl_Client_1	:	REAL:=250		;
		
		r_Water_PumpCIP_1		:	INT:=100	;
		r_Water_PumpClient_1	:	INT:=100	;
		
	*)


END_STRUCT
END_TYPE

// ---- 03 Project/23 CIP/str_ConcParam.TcDUT
TYPE str_ConcParam :
	//to be deletd
STRUCT
	
    r_Temper_1			:	REAL:=65	;//temperature set point for local client in celsius
	r_Flow_Pmp1_1		:	REAL:=180	;
	r_Flow_Pmp1_2		:	REAL:=180	;
	r_Pressure_Pmp1_1	:	REAL:=0.5	;
	r_Concentration_1	:	REAL:=0.3	;//concentration in percents
	t_Measure_Delay_1	:	INT:=60		;//measurment delay in seconds
END_STRUCT
END_TYPE

// ---- 03 Project/23 CIP/ST_CIP_Request.TcDUT
TYPE ST_CIP_Request :
STRUCT
	eType	: E_CIP_Type;
	eClient	: E_CIP_Usage;
	nClientId	: INT;					//1..30, 0 for eLocal
	eClientType	: E_Anybus_ClientType;	//eExternal only
	eStartState	: E_Element_State_Long;	//eExternal only: first stage, by the GAD wash type

END_STRUCT
END_TYPE

// ---- 03 Project/31 AnybusCommunication/E_Anybus_Alarm.TcDUT
{attribute 'qualified_only'}
{attribute 'to_string'}
//Interface alarm codes 1..99; CIP process alarm codes start from 100 (same word 6)
TYPE E_Anybus_Alarm :
(
	eNone				:= 0,
	eFieldbus			:= 1,	// gateway EtherCAT slave not in OP
	eAliveLost			:= 2,	// Siemens ALIVE does not toggle
	eRequestConflict	:= 3,	// REQUEST ON and REQUEST OFF together
	eInvalidClient		:= 4,	// CLIENT ID out of 1..30 with REQUEST ON
	eInvalidRecipe		:= 5,	// RECIPE TYPE not defined with REQUEST ON
	eInvalidClientType	:= 6	// CLIENT TYPE not defined with REQUEST ON
);
END_TYPE

// ---- 03 Project/31 AnybusCommunication/E_Anybus_ClientType.TcDUT
{attribute 'qualified_only'}
{attribute 'to_string'}
TYPE E_Anybus_ClientType :
(
	eNone	:= 0,	// not selected
	ePipe	:= 1,	// no spray ball
	eTank	:= 2	// always with a spray ball, decided 01.11.2026
);
END_TYPE

// ---- 03 Project/31 AnybusCommunication/E_Anybus_Media.TcDUT
{attribute 'qualified_only'}
{attribute 'to_string'}
TYPE E_Anybus_Media :
(
	eNone				:= 0,	// no sending
	eFirstWater			:= 1,	// pre-rinse, T93 recycle water
	eSoda				:= 2,	// detergent, T92
	eIntermediateWater	:= 3,	// T94 water
	eDisinfection		:= 4,	// T91
	eLastWater			:= 5	// final rinse, T94 water
);
END_TYPE

// ---- 03 Project/31 AnybusCommunication/E_Anybus_RecipeType.TcDUT
{attribute 'qualified_only'}
{attribute 'to_string'}
TYPE E_Anybus_RecipeType :
(
	eNone			:= 0,	// not selected
	eFlushOnly				:= 1,	// CIP1
	eDetergent				:= 2,	// CIP1, CIP2, CIP3
	eDetergentOnly			:= 3,	// CIP2, CIP3
	eDisinfectionOnly		:= 4,	// CIP4, CIP5
	eDetergentDisinfection	:= 5,	// CIP2 .. CIP5
	eFull					:= 6	// CIP1 .. CIP5, codes proposed to GAD 02.11.2026
);
END_TYPE

// ---- 03 Project/31 AnybusCommunication/E_Anybus_Request.TcDUT
{attribute 'qualified_only'}
{attribute 'to_string'}
TYPE E_Anybus_Request :
(
	eNone		:= 0,	// ON=0, OFF=0: before start - idle, during CIP - pause
	eOn			:= 1,	// ON=1, OFF=0: run
	eOff		:= 2,	// ON=0, OFF=1: full stop
	eConflict	:= 3	// ON=1, OFF=1: not defined, treated as stop
);
END_TYPE

// ---- 03 Project/31 AnybusCommunication/E_Sim_Fault.TcDUT
{attribute 'qualified_only'}
{attribute 'to_string'}
TYPE E_Sim_Fault :
(
	eNone			:= 0,
	ePause			:= 1,	// PAUSE from the plant
	eInletOff		:= 2,	// INLET PUMP ENABLE = 0
	eRequestDrop	:= 3,	// REQUEST ON lost, no REQUEST OFF
	eRequestOff		:= 4,	// REQUEST OFF in the middle of the wash
	eConflict		:= 5,	// REQUEST ON and OFF together
	eAliveStop		:= 6,	// ALIVE does not toggle
	eCable			:= 7,	// all data 0, like a pulled cable
	eBadClient		:= 8,	// CLIENT ID out of range
	eBadRecipe		:= 9,	// RECIPE TYPE out of range
	eBadType		:= 10,	// CLIENT TYPE out of range
	eNextUnstable	:= 11,	// NEXT CLIENT changes every second
	eNoClientEmpty	:= 12,	// CLIENT EMPTY is not answered
	eNoSprinkler	:= 13,	// Sprinkler State is not answered
	eReadyOff		:= 14	// plant READY = 0
);
END_TYPE

// ---- 03 Project/31 AnybusCommunication/E_Sim_Mode.TcDUT
{attribute 'qualified_only'}
{attribute 'to_string'}
TYPE E_Sim_Mode :
(
	eManual	:= 0,	// every signal is set by hand
	eAuto	:= 1,	// one wash cycle
	eQueue	:= 2	// clients of arQueue one after another
);
END_TYPE

// ---- 03 Project/31 AnybusCommunication/ST_Sim_Client.TcDUT
//One client of the Siemens simulator
TYPE ST_Sim_Client :
STRUCT
	nClient	: INT;					//0 = empty position
	eRecipe	: E_Anybus_RecipeType;
	eType	: E_Anybus_ClientType;
END_STRUCT
END_TYPE

// ---- 03 Project/31 AnybusCommunication/ST_Anybus_Inputs.TcDUT
//Siemens -> CIP, decoded from gIO.Anybus_Inputs_Raw
TYPE ST_Anybus_Inputs :
STRUCT
	//Word 0, byte 0
	bAlarm				: BOOL;	//0.0 plant alarm that stops CIP
	bReady				: BOOL;	//0.1 plant ready
	bRequestOn			: BOOL;	//0.2 start sending, held TRUE until REQUEST OFF
	bRequestOff			: BOOL;	//0.3 full stop
	bInletPumpEnable	: BOOL;	//0.4 enables the CIP sending pump
	bPause				: BOOL;	//0.5 pause from plant
	bClientEmpty		: BOOL;	//0.6 client is emptied (agreed 28.10.2026)
	bAlive				: BOOL;	//0.7 toggles 0.5 s / 0.5 s
	bSprinklerState		: BOOL;	//1.0 spray ball route is ready (proposal)

	nClientId			: INT;					//word 1, 1..30
	eRecipeType			: E_Anybus_RecipeType;	//word 2
	eClientType			: E_Anybus_ClientType;	//word 3
	nNextClient			: INT;					//word 4, 0 = none
	eNextRecipe			: E_Anybus_RecipeType;	//word 5
	eNextClientType		: E_Anybus_ClientType;	//word 6 (CIP proposal)
END_STRUCT
END_TYPE

// ---- 03 Project/31 AnybusCommunication/ST_Anybus_Outputs.TcDUT
//CIP -> Siemens, encoded to gIO.Anybus_Outputs_Raw
TYPE ST_Anybus_Outputs :
STRUCT
	//Word 0, byte 0
	bAlarm				: BOOL;	//0.0 CIP alarm
	bReady				: BOOL;	//0.1 solution for the next client is prepared
	bWorking			: BOOL;	//0.2 CIP in progress
	bFinish				: BOOL;	//0.3 CIP finished
	bEmptyingClient		: BOOL;	//0.4 client must be emptied between media
	bSendingPump		: BOOL;	//0.5 sending pump is running
	bPause				: BOOL;	//0.6 CIP is paused
	bAlive				: BOOL;	//0.7 generated by FB_Anybus_Interface, value shown in fbAnybus.stOut
	bSprinklerRequest	: BOOL;	//1.0 level: 1 = spray ball needed, 0 = pipe (Vadim 02.11.2026, address not agreed with GAD)

	eActualMedia		: E_Anybus_Media;		//word 1
	nRecipeProgress		: DINT;					//words 2-3, setpoint of the current stage
	nActualProgress		: DINT;					//words 4-5, actual value of the current stage
	nAlarmCode			: INT;					//word 6, 0 = no alarm, CIP process codes from 100 (proposal)
	nProgressUnit		: INT;					//word 7, 1 = seconds, 2 = litres (proposal)
	nActiveClient		: INT;					//word 8, echo of the client in CIP (proposal)
	eActiveRecipe		: E_Anybus_RecipeType;	//word 9, echo of the recipe in CIP (proposal)
	nFlowRateSet		: INT;					//word 10, required flow rate (proposal)
	nFlowRateActual		: INT;					//word 11, actual flow rate (proposal)
END_STRUCT
END_TYPE

// ---- 00 Library/00-General/TimeAndDate/GVL_Time_12.TcGVL

VAR_GLOBAL
		(*----------------> Real Time Clock <------------------*)

	dtRealTime								:DATE_AND_TIME;
	sRealTime								:STRING[22];
	stSystemTime							:TimeStruct;
	stSystemTime_Empty						:TimeStruct;
	sDateShort								:STRING[20];	(*	YYMMDD	*)
	
(*..........................................................................System TIME.....................................................................................*)
	sTime					: STRING[20];
	sDate					: STRING[20];
	sDateTime				: STRING[60];
	sTimeWithMicroSec		: STRING[40];

END_VAR

// ---- 00 Library/04 Recipe/GVL_Recipe.TcGVL
//{attribute 'qualified_only'}
VAR_GLOBAL CONSTANT	
	C_Max_RecipeFileNum				: INT:=100;
	C_Max_Recipe_List				: INT:=E_Recipe_Name.R_Piston_Settings;

END_VAR

VAR_GLOBAL 
	fbRecipe					: ARRAY [1..C_Max_Recipe_List] OF FB_Recipe;
	stRecipe					: ARRAY [1..C_Max_Recipe_List] OF ST_Recipe;

	ar_RecipesLoadDefault			: ARRAY [1..E_Recipe_Name.R_Piston_Settings] OF BOOL;
	ar_RecipesStoragePath			: ARRAY [1..E_Recipe_Name.R_Piston_Settings] OF STRING(80);;	
	
END_VAR

VAR_GLOBAL PERSISTENT
	eRecipeRootFolder: E_Recipe_Root_Folder:=E_Recipe_Root_Folder.PLC;
	ar_RecipesStoragePath_Root			: ARRAY [0..4] OF STRING:=[	
	(*PLC*)			'C:\Recipe',
	(*Develop_1*)	'C:\Users\admin\Source\Repos\RM003_PLC\Recipes',
	(*Develop_2*)	'C:\Users\admin\Source\Repos\RM003_PLC\RM003_PLC\Recipe',
	(*Develop_3*)	'C:\Users\dell\source\repos\KFM001_Hyper\Recipes',
	(*Develop_4*)	'\Hard Disk\ftp\Recipe'
	];		
	
	ar_RecipesStoragePath_Folder			: ARRAY [1..C_Max_Recipe_List] OF STRING;			
	
END_VAR

// ---- 00 Library/04-Messages/GVL_CycleMessages.TcGVL
//{attribute 'qualified_only'}
VAR_GLOBAL
	Buffer_Act_Message				:ARRAY[1..C_Max_Buffer_Act_list] OF stMessageFormat;
	Buffer_Act_Warning				:ARRAY[1..C_Max_Buffer_Act_list] OF stMessageFormat;
	Buffer_Act_History				:ARRAY[1..C_Max_Buffer_Act_list] OF stMessageFormat;
	Buffer_Search_Messages			:ARRAY[1..1000] OF stMessageFormat;
	Buffer_Act_Display				:ARRAY[1..20] 	OF stMessageFormat;

	fbPrintErrMessageByID			:FB_PrintErrMessageByID;	

	s_Error_BitmapID	       		:STRING;
	
	ar_ErrorActive					:ARRAY[1..C_Max_ErrorList] 	OF BOOL;	
	

	
END_VAR
VAR_GLOBAL CONSTANT
	C_Max_ErrorList: INT:=200;
	C_Max_Buffer_Act_list: INT:=100;

END_VAR

// ---- 00 Library/05 Safety/GVL_Safety.TcGVL
VAR_GLOBAL
	//bStateSafe						:BOOL:=TRUE; // FALSE
	
	bES_Bypass						:BOOL:=FALSE;

	 // FALSE
	bES_Relay						:BOOL; 
	bES_Relay_FB					:BOOL; 

	//stSafetyIn			AT %I* 		:ST_SafeIn;
	//stSafetyOut			AT %Q* 		:ST_SafeOut;

	bES_PB							:ARRAY[1..12] 	OF ST_ES_PB;
	bInterlock						:ARRAY[1..12] 	OF BOOL;
	bDoorLocked						:ARRAY[1..12] 	OF BOOL;
	bInterlockZone		AT %I*	 	:ARRAY[1..4] 	OF BOOL;
	bIntZoneLocked					:ARRAY[1..4] 	OF BOOL;
	bIntZoneBypass			 		:ARRAY[1..4] 	OF BOOL;
	bReq_LockZone					:ARRAY[1..4] 	OF BOOL;
	
	sBitmap_ESButton		     	:STRING; //for visualization
	stBitMap                		:STRING; //for HMI
 
    sInterlocksZone1                 :STRING; 
    sInterlocksZone2                 :STRING; 
    sInterlocksZone3                 :STRING; 
   	sInterlocksZone4                 :STRING; 	
END_VAR

// ---- 00 Library/11 HMI/g_HMI.TcGVL
//{attribute 'qualified_only'}
VAR_GLOBAL
	eLed_Color: E_Led_Color;
	
	eProcessControl_Name	: E_ProcessControl_Name	;
	
	eCIP_DashStage			: E_CIP_DashStage	;
	eCIP_DashStage_actual	: E_CIP_DashStage_List;
	sCIP_DashStage_actual	: STRING	;

	arCIP_DashStage_list	: ARRAY[0..E_CIP_DashStage_List.eLast] OF E_CIP_DashStage;
	arCIP_DashStage_string	: ARRAY[0..E_CIP_DashStage_List.eLast] OF STRING;
	arCIP_DashStage_MixProof: ARRAY[1..8] OF ST_MixProof_state;

	
	stT91_Sens		: ST_Tank_Level;
	stT92_Sens		: ST_Tank_Level;
	stT93_Sens		: ST_Tank_Level;
	stT94_Sens		: ST_Tank_Level;
	stT1_Sens		: ST_Tank_Level;
	stT2_Sens		: ST_Tank_Level;
	stT3_Sens		: ST_Tank_Level;
	stT4_Sens		: ST_Tank_Level;
END_VAR

// ---- 01 Instance/00-General/Global_Constant.TcGVL
//{attribute 'qualified_only'}
VAR_GLOBAL CONSTANT
	//C_Max_ErrorList				: INT:=200;
	//C_Max_Pistons				: INT:=7;
	//C_Max_MotorsAC				: INT:=6;
	//C_Max_Measure				: INT:=15;
END_VAR

// ---- 01 Instance/00-General/Global_Persistent.TcGVL
//{attribute 'Tc2GvlVarNames'}
VAR_GLOBAL PERSISTENT
	Errors: DINT;
	SetSlaveToOP_ON     : BOOL:=TRUE;
	bEnableAutoResetEncoder: BOOL:=TRUE;
END_VAR

// ---- 01 Instance/00-General/VersionDescription.TcGVL
//{attribute 'qualified_only'}
VAR_GLOBAL CONSTANT
	ProgramVersion: 			STRING	:=	'V0.1.0.0';			(*	Product . Major . Revision . Build	*)
(*
V0.1.0.0 	- Start version menager.
				- ...

*)	
END_VAR

// ---- 01 Instance/01 Piston/g_Piston.TcGVL
//{attribute 'qualified_only'}
VAR_GLOBAL	
	fbPis			: ARRAY[0..E_Pis_Name.last] OF FB_Piston;
	stPis			: ARRAY[0..E_Pis_Name.last] OF ST_Piston;
	arPisName		: ARRAY[0..E_Pis_Name.last] OF ST_Piston_SelectionList;
	

	iPis_sel		: INT:=1;
	
	arPisNameList	: ARRAY[0..E_Pis_Name.last] OF STRING(12);
	ePisNameList	: E_Pis_Name;

	fbPis_U_L		: ARRAY[0..E_Pis_Name.last] OF FB_Piston_U_L;
	stPis_U_L		: ARRAY[0..E_Pis_Name.last] OF ST_Piston_U_L;

	
END_VAR

VAR_GLOBAL PERSISTENT
	stPisSetting	: ARRAY[0..E_Pis_Name.last] OF ST_Piston_Setting_Param;
END_VAR

VAR_GLOBAL CONSTANT
	C_MAX_Pistons		: INT:=E_Pis_Name.last;
	//C_MAX_Pistons_Exist	: INT:=51;	
END_VAR

// ---- 01 Instance/02 Pump/g_Pump.TcGVL
//{attribute 'qualified_only'}
VAR_GLOBAL
	fbPump			: ARRAY[0..E_Pump_List.last] OF FB_Pump	;
	arr_st_Pump		: ARRAY[0..E_Pump_List.last] OF ST_Pump	;
	
	fbDosingPP1002: FB_DosingPump; //Detergent
	fbDosingPP1003: FB_DosingPump; //DisInfection

END_VAR

// ---- 01 Instance/03 SFC/g_SFC.TcGVL
{attribute 'qualified_only'}
VAR_GLOBAL
	fbSFC_Temp1: FB_SFC_Template;
END_VAR

// ---- 01 Instance/04-Messages/Error_List.TcGVL
VAR_GLOBAL

END_VAR

VAR_GLOBAL CONSTANT
	
	ar_ErrorList					:ARRAY[1..C_Max_ErrorList,0..2] 	OF STRING[80]:= [
(*	Error ID				Error ID		Error Message_ _ _ _ _ _  _ _ _ _ _ _ _ _ _ _ _ _ _ _ _ _ _ _ _ _*)
		(*8888888888888888888888888888888888888888888*)					


		                  (************************************ General *****************************************)

'000x000xPUZ',   'Message',   'Pause requested',

'000x000x999',	  'Error',	  'General Error',
'000x000x777',	  'Error',	  'EtherCAT Com Fault - Chack Hardware Configuration',
'777x777x777',	  'Error',	  'Loading Carrier Is Ready to move without Top Plate - logic conflict',

'SMTx000x001',	  'Error',	  'Servo motor General Error',
'SMTx000x002',	  'Error',	  'Servo motor Power Not OK',

'050x000x001',  'Error',   'Air Pressure Too Low',
'050x000x002',  'Message', 'Production Finished',
'050x000x003',  'Error',   'Not able to change to Semi or Auto mode befor General initialization done',
'050x000x004',  'Error',   'Unknown carrier status detected',
'050x000x005',  'Error',   'Suction Tank Over Flow',
'050x000x300',	'Warning',	'Manual mode request rejected - first pause automation',
'050x000x301',	'Warning',	'Semi mode request rejected - first pause automation',
'050x000x302',	'Warning',	'Auto mode request rejected - first pause automation',
'050x000x303',	'Warning',	'Manual mode request rejected - Pistion not in last auto pisition',
'050x000x304',	'Warning',	'Semi mode request rejected - Pistion not in last auto pisition',
'050x000x305',	'Warning',	'Auto mode request rejected - Pistion not in last auto pisition',
'050x000x306',	'Warning',	'Semi/Auto mode request rejected - automation lock failed',

'050x000x350',	'Warning',	'Semi/Auto mode request rejected - initialize all system first',
'050x000x351',	'Warning',	'Interlock Paused Operation',

    (*CIP Tanks Overweight and overflow*)
'101x000x000',   'Warning',      'CIP Tanks Overweight >> 1500 liter',
'101x000x001',   'Warning',      'CIP Tank T91 overflow',
'101x000x002',   'Warning',      'CIP Tank T92 overflow',
'101x000x003',   'Warning',      'CIP Tank T93 overflow',
'101x000x004',   'Warning',      'CIP Tank T94 overflow',

	(*CIP Tanks concentration delution*)
'101x000x101',   'Warning',      'CIP - Detergent concentration delution requered',
'101x000x102',   'Warning',      'CIP - Detergent concentration delution limited by tank max volume',
'101x000x103',   'Error',      	 'CIP - Detergent concentration delution limited by tank max volume',

'101x000x111',   'Warning',      'CIP - DisInfection concentration delution requered',
'101x000x112',   'Warning',      'CIP - DisInfection concentration delution limited by tank max volume',
'101x000x113',   'Error',      	 'CIP - DisInfection concentration delution limited by tank max volume',

	(*Pumps*)
'P1001x001',   	'Error',      'Motor driver is not ready at run',
'P3001x001',   	'Error',      'Motor driver is not ready at run',
'P3002x001',   	'Error',      'Motor driver is not ready at run',
'AG3001x001',   'Error',      'Motor driver is not ready at run',
'AG3002x001',   'Error',      'Motor driver is not ready at run',
'P4001x001',   	'Error',      'Motor driver is not ready at run',
'P4002x001',   	'Error',      'Motor driver is not ready at run',
'AG4001x001',   'Error',      'Motor driver is not ready at run',
'AG4002x001',   'Error',      'Motor driver is not ready at run',
'TB0001x001',   'Error',      'Motor driver is not ready at run',

'P1001x002',   	'Warning',      'Motor speed feedback lag monitoring',
'P3001x002',   	'Warning',      'Motor speed feedback lag monitoring',
'P3002x002',   	'Warning',      'Motor speed feedback lag monitoring',
'AG3001x002',   'Warning',      'Motor speed feedback lag monitoring',
'AG3002x002',   'Warning',      'Motor speed feedback lag monitoring',
'P4001x002',   	'Warning',      'Motor speed feedback lag monitoring',
'P4002x002',   	'Warning',      'Motor speed feedback lag monitoring',
'AG4001x002',   'Warning',      'Motor speed feedback lag monitoring',
'AG4002x002',   'Warning',      'Motor speed feedback lag monitoring',
'TB0001x002',   'Warning',      'Motor speed feedback lag monitoring',

'P1001x003',   	'Warning',      'Motor driver is not ready',
'P3001x003',   	'Warning',      'Motor driver is not ready',
'P3002x003',   	'Warning',      'Motor driver is not ready',
'AG3001x003',   'Warning',      'Motor driver is not ready',
'AG3002x003',   'Warning',      'Motor driver is not ready',
'P4001x003',   	'Warning',      'Motor driver is not ready',
'P4002x003',   	'Warning',      'Motor driver is not ready',
'AG4001x003',   'Warning',      'Motor driver is not ready',
'AG4002x003',   'Warning',      'Motor driver is not ready',
'TB0001x003',   'Warning',      'Motor driver is not ready',


// Pump Pressure is dangerously high
'P1001x004',   	'Error',      'Pump Pressure is dangerously high',
'P3001x004',   	'Error',      'Pump Pressure is dangerously high',
'P3002x004',   	'Error',      'Pump Pressure is dangerously high',
'P4001x004',   	'Error',      'Pump Pressure is dangerously high',
'P4002x004',   	'Error',      'Pump Pressure is dangerously high',
// Pump Pressure is above normal
'P1001x005',   	'Warning',      'Pump Pressure is above normal',
'P3001x005',   	'Warning',      'Pump Pressure is above normal',
'P3002x005',   	'Warning',      'Pump Pressure is above normal',
'P4001x005',   	'Warning',      'Pump Pressure is above normal',
'P4002x005',   	'Warning',      'Pump Pressure is above normal',
// Pump Pressure is below normal
'P1001x006',   	'Warning',      'Pump Pressure is below normal',
'P3001x006',   	'Warning',      'Pump Pressure is below normal',
'P3002x006',   	'Warning',      'Pump Pressure is below normal',
'P4001x006',   	'Warning',      'Pump Pressure is below normal',
'P4002x006',   	'Warning',      'Pump Pressure is below normal',
// Pump Pressure is critically low
'P1001x007',   	'Error',      'Pump Pressure is critically low',
'P3001x007',   	'Error',      'Pump Pressure is critically low',
'P3002x007',   	'Error',      'Pump Pressure is critically low',
'P4001x007',   	'Error',      'Pump Pressure is critically low',
'P4002x007',   	'Error',      'Pump Pressure is critically low',

//Manual mode active
'P1001x008',   	'Warning',      'Motor manual mode active',
'P3001x008',   	'Warning',      'Motor manual mode active',
'P3002x008',   	'Warning',      'Motor manual mode active',
'AG3001x008',   'Warning',      'Motor manual mode active',
'AG3002x008',   'Warning',      'Motor manual mode active',
'P4001x008',   	'Warning',      'Motor manual mode active',
'P4002x008',   	'Warning',      'Motor manual mode active',
'AG4001x008',   'Warning',      'Motor manual mode active',
'AG4002x008',   'Warning',      'Motor manual mode active',
'TB0001x008',   'Warning',      'Motor manual mode active',

'101x001x001',   'Error',      'Message num 1, non cyclic',
'101x001x002',   'Message',    'Waiting for Operator to Start Single Cycle',
'101x001x003',   'Error',      'Stepper did not found paper',
'101x001x004',   'Warning',    'Gripper Cycle without moving Stepper',
'101x001x005',   'Error',      'Multiple Gripper Cycles without moving Stepper',
'101x001x006',   'Warning',    'Paper Ended in Run mode',
'101x001x007',   'Warning',    'Paper Stacker Empty on Paper Check',
'101x001x008',   'Error',      'Paper Stacker Column hight diference exceeds allowed limit',
'101x001x009',   'Warning',     'System is waiting for Resume or Play activation from Operator',
'101x001x010',   'Error',     	'Gripper Encoder is over 25000 the limit',
'101x001x011',   'Warning',     'Stepper stopped, did not found papper',

 (*Tanks Interlock*)
'101x002xT91',   'Error',      'CIP Tank T91 in not locked',
'101x002xT92',   'Error',      'CIP Tank T92 in not locked',
'101x002xT93',   'Error',      'CIP Tank T93 in not locked',
'101x002xT94',   'Error',      'CIP Tank T94 in not locked',

'101x002xT01',   'Warning',      'Marinade Tank T01 in not locked',
'101x002xT02',   'Warning',      'Marinade Tank T02 in not locked',

'101x002xT03',   'Error',      'Color Tank T03 in not locked',
'101x002xT04',   'Error',      'Color Tank T04 in not locked',

